	xInit			: BOOL;
	diPosPrev		: DINT;
	diTargetPrev	: DINT;
	diMoveStart		: DINT;

	xDirRev			: BOOL;
	xNewMove		: BOOL;
	xMoveWanted		: BOOL;
	xBrakeOpen		: BOOL;
	xMoving			: BOOL;
	xRunPrev		: BOOL;

	diStopAccum		: DINT;
	xCoasting		: BOOL;

	rtrgGo			: R_TRIG;
	rtrgReset		: R_TRIG;
	rtrgSetAccum	: R_TRIG;

	tofBrake		: TOF;
	tonBrakeOpen	: TON;
	tonGrace		: TON;
	tonStall		: TON;
	tonRest			: TON;
	tonDrvAck		: TON;

	diStallRef		: DINT;
	xStallReset		: BOOL;
	xStallArmed		: BOOL;

END_VAR

// =============================================================
// ENKODER -> PRZYROST ZE ZNAKIEM
// =============================================================
//
// Surowa wartosc moze byc wieksza niz jeden obrot, wiec
// sprowadzamy ja modulo. MOD na ujemnej daje w ST wynik ujemny,
// dlatego domykamy recznie.

diPos := diRawPos MOD 65536;

IF diPos < 0 THEN
	diPos := diPos + 65536;
END_IF


IF NOT xInit THEN
	xInit        := TRUE;
	diPosPrev    := diPos;
	diStallRef   := diPos;
	diTargetPrev := diTargetAbs;
END_IF


// Skok wiekszy niz pol obrotu nie jest ruchem - to licznik
// przekrecil sie przez zero. Prostujemy go i liczymy przejscie.

diStep := diPos - diPosPrev;

IF diStep > 32768 THEN
	diStep  := diStep - 65536;
	diTurns := diTurns - 1;
END_IF

IF diStep < -32768 THEN
	diStep  := diStep + 65536;
	diTurns := diTurns + 1;
END_IF

diPosPrev := diPos;


// =============================================================
// POZYCJA NARASTAJACA
// =============================================================
//
// Tu przestaje istniec problem przekrecania sie enkodera.
// diAccum jest zwykla liczba impulsow od punktu odniesienia
// i rosnie miedzy obrotami bez zadnego zawijania.

diAccum := diAccum + diStep;


// Punkt odniesienia ustawiany z zewnatrz, raz na cykl
rtrgSetAccum(CLK := xSetAccum);

IF rtrgSetAccum.Q THEN
	diAccum     := diSetAccumTo;
	diMoveStart := diSetAccumTo;
	xInPos      := TRUE;

	// Pomiar dojazdu musi przejsc przez ten skok sucha stopa.
	// diCoast liczy sie jako roznica na skali narastajacej,
	// wiec przestawienie punktu odniesienia bez tego wygladalo
	// by jak dojazd o caly obrot.
	diStopAccum := diSetAccumTo;
	xCoasting   := FALSE;
END_IF


// =============================================================
// NOWY RUCH
// =============================================================
//
// Nowy ruch to podanie zadania albo zmiana celu. diTargetAbs
// ma byc STALA w obrebie kroku - inaczej kazdy cykl wygladalby
// jak nowy ruch.

rtrgGo(CLK := xGoTo AND xEnable);

xNewMove := rtrgGo.Q OR (diTargetAbs <> diTargetPrev);
diTargetPrev := diTargetAbs;

IF xNewMove THEN
	diMoveStart := diAccum;
	xInPos      := FALSE;
	diStallRef  := diPos;
END_IF


// =============================================================
// UCHYB I KONIEC RUCHU
// =============================================================
//
// Zwykle odejmowanie, bez modulo. Uchyb ujemny znaczy "cel juz
// przejechany" i konczy ruch NATYCHMIAST - to jest dokladnie
// ten przypadek, w ktorym stara wersja wysylala os na dodatkowy
// pelen obrot.
//
// xInPos jest zatrzaskiem: osuniecie sie wozka po zacisnieciu
// hamulca nie ma prawa odwolac zaliczonego kroku.

diRemain := diTargetAbs - diAccum;
diMoved  := diAccum - diMoveStart;

IF diRemain <= diStopLead THEN
	xInPos := TRUE;
END_IF


// =============================================================
// RUCH I HAMULEC
// =============================================================
//
// Hamulec idzie za ZADANIEM ruchu, falownik dostaje komende
// tBrakeReleaseLead pozniej. Przy zerze - jednoczesnie.

xJogging := xEnable AND (xJogFwd XOR xJogRev);

xMoveWanted := xEnable AND NOT xStall AND (xJogging OR (xGoTo AND NOT xInPos));

// W cyklu korba jedzie WYLACZNIE do przodu. Kierunek wymuszamy
// co cykl, zeby ten z jazdy recznej w tyl nie mogl przezyc.
xDirRev := FALSE;

IF xJogging THEN
	xDirRev := xJogRev;
END_IF


tofBrake(IN := xMoveWanted, PT := tBrakeHold);
xBrakeRelease := tofBrake.Q;

tonBrakeOpen(IN := xMoveWanted AND xBrakeRelease, PT := tBrakeReleaseLead);

// Warunek na zero jawny - nie opieramy sie na tym, jak TON
// zachowa sie przy PT = 0. Blad w te strone dalby os, ktora
// nigdy nie rusza, i nic by tego nie powiedzialo.
xBrakeOpen := tonBrakeOpen.Q OR (tBrakeReleaseLead = T#0S);

xBrakeWait := xMoveWanted AND NOT xBrakeOpen;

xMoving := xMoveWanted AND xBrakeRelease AND xBrakeOpen;

xRunReq := xMoving;
xRev    := xDirRev;


// =============================================================
// POMIAR DOJAZDU
// =============================================================

IF xRunPrev AND NOT xRunReq THEN
	diStopAccum := diAccum;
	xCoasting   := TRUE;
END_IF

xRunPrev := xRunReq;

IF xCoasting THEN
	diCoast := diAccum - diStopAccum;
END_IF

tonRest(IN := ABS(diStep) < diStallMin, PT := tRest);
xAtRest := tonRest.Q;

IF xAtRest THEN
	xCoasting := FALSE;
END_IF


// =============================================================
// CZUWAK RUCHU
// =============================================================
//
// Uzbrojony dopiero po tStallGrace od startu - hamulec musi
// odpuscic, a silnik rozbiec sie rampa.

tonGrace(IN := xRunReq, PT := tStallGrace);
xStallArmed := tonGrace.Q;

xStallReset := (ABS(diAccum - diStallRef) > diStallMin)
               OR NOT xStallArmed OR xNewMove;

IF xStallReset THEN
	diStallRef := diAccum;
END_IF

tonStall(IN := xStallArmed AND NOT xStallReset, PT := tStall);

IF tonStall.Q THEN
	xStall := TRUE;
END_IF


// -------------------------------------------------------------
// POTWIERDZENIE PRACY Z FALOWNIKA
// -------------------------------------------------------------
//
// Osobny, szybszy czuwak. Zadanie poszlo, hamulec zdjety,
// a falownik nie melduje pracy - nic nie trzyma wozka i nie ma
// na co czekac pelnych pieciu sekund.

tonDrvAck(IN := xRunReq AND NOT xDrvRunning, PT := tDrvAck);

IF tonDrvAck.Q THEN
	xNoDrvAck := TRUE;
	xStall    := TRUE;
END_IF


rtrgReset(CLK := xReset);

IF rtrgReset.Q OR NOT xEnable THEN
	xStall     := FALSE;
	xNoDrvAck  := FALSE;
	diStallRef := diAccum;
END_IF

END_FUNCTION_BLOCK

// ---- POUs/POUs/FB/FB_NordSK550PP.TcPOU
FUNCTION_BLOCK FB_NordSK550PP
// =============================================================
// NORDAC PRO SK 550P
// EtherCAT, profil NORD wg BU 2300 (NIE CiA 402)
// =============================================================
//
// FB nie wykonuje ZADNYCH operacji na predkosci.
// Zadanie jest podawane na stale, sterowanie odbywa sie
// wylacznie bitami ControlWord. Rozpedzanie i hamowanie
// realizuje falownik parametrami P102 / P103 / P108.
//
// Sterowanie przez metody:
//   M_Start(lrFreq, xReverse)   - zadanie + bit startu
//   M_Stop()                    - zdjecie bitu startu
//   M_Reset()                   - kasowanie bledow
//   M_SetFrequency(lrFreq)      - zmiana zadania
//
// Metody wywolywac PRZED cyklicznym wywolaniem instancji.
VAR_INPUT

	// P105 Maksymalna czestotliwosc falownika [Hz].
	// MUSI byc rowna P105 w falowniku - inaczej skalowanie
	// zadania jest bledne i naped dostaje inna czestotliwosc
	// niz zadana.
	lrFmax			: LREAL := 50.0;

	// TRUE = STO zwolnione, lancuch bezpieczenstwa OK
	xSafetyOK		: BOOL;

	// TRUE = komunikacja EtherCAT sprawna
	xEtherCAT_OK	: BOOL;

	// Dane procesowe z falownika
	stIn			: ST_NordSK550P_In;

END_VAR
VAR_OUTPUT

	// Dane procesowe do falownika
	stOut			: ST_NordSK550P_Out;


	// =========================================================
	// STATUS
	// =========================================================

	eState			: E_NordSK550P_State;

	xReadyToSwitchOn	: BOOL;
	xOperationEnabled	: BOOL;
	xSwitchOnInhibit	: BOOL;

	xRunning		: BOOL;
	xStopped		: BOOL;

	xFault			: BOOL;
	xWarning		: BOOL;
	xBusControl		: BOOL;

	xError			: BOOL;
	xCommError		: BOOL;


	// =========================================================
	// VALUES
	// =========================================================

	// Zadanie wysylane do falownika [Hz]
	lrFreqSetpoint	: LREAL;

	// Czestotliwosc rzeczywista z falownika [Hz]
	lrFreqActual	: LREAL;


	// =========================================================
	// DIAGNOSTICS
	// =========================================================

	wStatusWord		: UINT;
	wControlWord	: UINT;

	byModeDisplay	: USINT;

	//  0 = blokada, 10 = gotowosc, 20 = praca
	nStep			: INT;

END_VAR
VAR

	// Zadania z metod
	xReqRun			: BOOL;
	xReqReset		: BOOL;
	xReqReverse		: BOOL;
	lrReqFreq		: LREAL;

	wStateBits		: UINT;
	iSetpoint		: INT;
	xBlocked		: BOOL;

	tonComm			: TON;
	tonReset		: TON;

END_VAR
VAR CONSTANT

	// Skalowanie NORD: 16384 (0x4000) = 100% = P105
	cFullScale		: LREAL := 16384.0;

	// Prog zera dla czestotliwosci rzeczywistej [Hz]
	cZeroActual		: LREAL := 0.5;

	// ControlWord wg BU 2300 rozdz. 6.3.1
	//   047E = "Shut down"        - bit 0 zdjety, falownik
	//                               hamuje wlasna rampa P103
	//   047F = "Enable operation" - bit 0 zalaczony
	//   0480 = potwierdzenie bledu (bit 7)
	cCW_Shutdown	: UINT := 16#047E;
	cCW_EnableOp	: UINT := 16#047F;
	cCW_AckFault	: UINT := 16#0480;

	cCW_DirFwd		: UINT := 16#0800;
	cCW_DirRev		: UINT := 16#1000;

END_VAR

// =============================================================
// FB_NordSK550PP
// NORDAC PRO SK 550P - profil NORD wg BU 2300
// =============================================================
//
// ZASADA: PLC nie dotyka predkosci.
//
// Zadanie czestotliwosci jest podawane na stale i nie jest
// zerowane przy zatrzymaniu. Start to zalaczenie bitu 0
// ControlWord, stop to jego zdjecie. Reszte - rozpedzanie
// po P102, hamowanie po P103, sposob wygaszania po P108
// i ewentualne dohamowanie pradem stalym po P559 - robi
// falownik.
//
// ControlWord (BU 2300 rozdz. 6.3.1):
//   bit 0  Ready for operation   <-- start / stop
//   bit 1  Voltage disable       (1 = kasuj blokade napiecia)
//   bit 2  Quick stop            (1 = kasuj quick stop)
//   bit 3  Enable operation
//   bit 4  Enable pulses
//   bit 5  Enable ramp
//   bit 6  Setpoint enabled
//   bit 7  Acknowledge error     (zbocze 0 -> 1)
//   bit 10 Control data valid    <-- BEZ NIEGO NAPED IGNORUJE DANE
//   bit 11 CW, bit 12 CCW
//
// StatusWord (rozdz. 6.3.2), bity 0..6:
//   0x31 Ready to switch-on   0x33 Switched on
//   0x37 Operation enabled    0x17 Quick stop active
//   bit 3 Fault               bit 6 Switch-on inhibit
//
// Zadanie i wartosc rzeczywista sa procentowe:
//   16384 (0x4000) = 100% = P105
//
// Nazwy pol diTargetVelocity / iVelocityDemand w ST_NordSK550P_*
// sa mylace - to NIE obroty, tylko czestotliwosc w skali
// procentowej. NIE zmieniac tych nazw: sa uzyte w linkach I/O
// w .tsproj dla wszystkich 19 napedow.


// =============================================================
// COPY INPUT DATA
// =============================================================

wStatusWord		:= stIn.wStatusWord;
byModeDisplay	:= stIn.byModeDisplay;

IF lrFmax > 0.0 THEN
	lrFreqActual := INT_TO_LREAL(stIn.iVelocityDemand) / cFullScale * lrFmax;
ELSE
	lrFreqActual := 0.0;
END_IF


// =============================================================
// COMMUNICATION WATCHDOG
// =============================================================

tonComm(IN := NOT xEtherCAT_OK, PT := T#500MS);
xCommError := tonComm.Q;


// =============================================================
// STATUSWORD DECODING
// =============================================================

xFault				:= (wStatusWord AND 16#0008) <> 0;
xWarning			:= (wStatusWord AND 16#0080) <> 0;
xSwitchOnInhibit	:= (wStatusWord AND 16#0040) <> 0;
xBusControl			:= (wStatusWord AND 16#0200) <> 0;

wStateBits := wStatusWord AND 16#007F;


IF xFault THEN

	IF (wStatusWord AND 16#000F) = 16#000F THEN
		eState := NORD_STATE_FAULT_REACTION_ACTIVE;
	ELSE
		eState := NORD_STATE_FAULT;
	END_IF

ELSIF xSwitchOnInhibit THEN
	eState := NORD_STATE_SWITCH_ON_DISABLED;

ELSIF wStateBits = 16#0031 THEN
	eState := NORD_STATE_READY_TO_SWITCH_ON;

ELSIF wStateBits = 16#0033 THEN
	eState := NORD_STATE_SWITCHED_ON;

ELSIF wStateBits = 16#0037 THEN
	eState := NORD_STATE_OPERATION_ENABLED;

ELSIF wStateBits = 16#0017 THEN
	eState := NORD_STATE_QUICK_STOP_ACTIVE;

ELSIF (wStatusWord AND 16#000F) = 0 THEN
	eState := NORD_STATE_NOT_READY;

ELSE
	eState := NORD_STATE_UNKNOWN;

END_IF


xReadyToSwitchOn	:= (eState = NORD_STATE_READY_TO_SWITCH_ON);
xOperationEnabled	:= (eState = NORD_STATE_OPERATION_ENABLED);


// =============================================================
// WARUNKI BLOKUJACE
// =============================================================

xBlocked := xFault OR xCommError OR NOT xSafetyOK;
xError   := xBlocked;


// =============================================================
// CONTROLWORD
// =============================================================
//
// Trzy stany, bez zadnej sekwencji posredniej. Przejscia
// wewnetrznej maszyny stanow falownika (Switch-on inhibit ->
// Ready to switch-on -> Switched on -> Operation enabled)
// realizuje sam falownik: 047E zawiera komende "Shut down",
// a 047F jednoczesnie "Switch on" i "Enable operation".

IF xBlocked THEN

	nStep := 0;

	// Zadanie ruchu kasujemy - po ustapieniu przyczyny naped
	// NIE moze ruszyc sam, operator musi wywolac M_Start.
	xReqRun := FALSE;

	wControlWord := 16#0000;

	// Kasowanie bledu: impuls na bicie 7
	IF xReqReset AND xSafetyOK AND NOT xCommError THEN
		wControlWord := cCW_AckFault;
	END_IF

ELSIF xReqRun THEN

	nStep := 20;
	wControlWord := cCW_EnableOp;

	// BLOKADA ZALACZENIA (Switch-on inhibit, bit 6 statusu).
	//
	// Ze stanu "Switch on disabled" falownik NIE wyjdzie na 047F.
	// Bit 0 musi zobaczyc zbocze, a zeby je zobaczyl, trzeba
	// najpierw wyslac Shutdown (047E). Trzymanie 047F w kolko
	// zostawia naped w blokadzie na zawsze: bez bledu, bez ruchu,
	// bez zadnego komunikatu - dokladnie to widzielismy na
	// napedzie 5 po przeciazeniu i na 8 po zaniku komunikacji.
	//
	// Dopoki falownik melduje blokade, wysylamy wiec 047E. Gdy
	// z niej wyjdzie, w nastepnym cyklu idzie juz 047F i naped
	// rusza sam, bez kasowania bledu i bez zdejmowania startu.
	IF xSwitchOnInhibit THEN
		nStep := 15;
		wControlWord := cCW_Shutdown;
	END_IF

ELSE

	nStep := 10;
	wControlWord := cCW_Shutdown;

END_IF


// =============================================================
// KIERUNEK
// =============================================================
//
// Zmiane kierunku w ruchu obsluguje falownik - przechodzi
// przez absolutna minimalna czestotliwosc P505.

IF wControlWord <> 16#0000 THEN

	IF xReqReverse THEN
		wControlWord := wControlWord OR cCW_DirRev;
	ELSE
		wControlWord := wControlWord OR cCW_DirFwd;
	END_IF

END_IF


// =============================================================
// IMPULS KASOWANIA BLEDU
// =============================================================
//
// Bit 7 musi zobaczyc zbocze 0 -> 1. Trzymamy go 200 ms,
// potem kasujemy zadanie, zeby kolejne M_Reset znowu
// wytworzylo zbocze.

tonReset(IN := xReqReset, PT := T#200MS);

IF tonReset.Q THEN
	xReqReset := FALSE;
END_IF


// =============================================================
// ZADANIE CZESTOTLIWOSCI
// =============================================================
//
// Podawane na stale. NIE zerujemy go przy zatrzymaniu -
// stop realizuje bit 0 ControlWord, a hamowanie falownik.

lrFreqSetpoint := lrReqFreq;

IF lrFreqSetpoint > lrFmax THEN
	lrFreqSetpoint := lrFmax;
END_IF

IF lrFreqSetpoint < 0.0 THEN
	lrFreqSetpoint := 0.0;
END_IF


IF lrFmax > 0.0 THEN
	iSetpoint := LREAL_TO_INT(lrFreqSetpoint / lrFmax * cFullScale);
ELSE
	iSetpoint := 0;
END_IF

IF iSetpoint > 16384 THEN
	iSetpoint := 16384;
END_IF

IF iSetpoint < 0 THEN
	iSetpoint := 0;
END_IF


// =============================================================
// WRITE OUTPUT PDO
// =============================================================
//
// byModeOfOperation nie jest zmapowany w .tsproj - falownik
// NORD nie uzywa obiektu 0x6060. Zostawiamy zero.

stOut.byModeOfOperation	:= 0;
stOut.wControlWord		:= wControlWord;
stOut.diTargetVelocity	:= iSetpoint;


// =============================================================
// STATUS WYJSCIOWY
// =============================================================

xRunning := xOperationEnabled AND NOT xBlocked;

xStopped := (ABS(lrFreqActual) <= cZeroActual);

METHOD M_Start : BOOL
VAR_INPUT
	// Zadana czestotliwosc [Hz]
	lrFreq		: LREAL;

	// FALSE = w prawo (CW), TRUE = w lewo (CCW)
	xReverse	: BOOL;
END_VAR
// Zadanie czestotliwosci + bit startu. Nic wiecej.
// Rozpedzanie realizuje falownik rampa P102.
//
// Zadanie jest zatrzaskiwane - obowiazuje az do M_Stop
// albo do wystapienia blokady (blad / STO / komunikacja).

lrReqFreq	:= lrFreq;
xReqReverse	:= xReverse;
xReqRun		:= TRUE;

M_Start := TRUE;
END_METHOD

METHOD M_Stop : BOOL
// Zdjecie bitu 0 ControlWord. Nic wiecej - zadanie
// czestotliwosci zostaje bez zmian.
//
// Falownik hamuje wlasna rampa P103, sposob wygaszania
// okresla P108, ewentualne dohamowanie pradem stalym P559.

xReqRun := FALSE;

M_Stop := TRUE;
END_METHOD

METHOD M_Reset : BOOL
// Kasowanie bledow falownika. FB wystawia impuls 200 ms
// na bicie 7 ControlWord (zbocze 0 -> 1 wg BU 2300).
//
// Dziala tylko wtedy, gdy przyczyna blokady ustapila:
// STO zwolnione i komunikacja sprawna.

xReqReset := TRUE;

M_Reset := TRUE;
END_METHOD

METHOD M_SetFrequency : BOOL
VAR_INPUT
	// Zadana czestotliwosc [Hz]
	lrFreq		: LREAL;
END_VAR
// Zmiana zadania. Falownik dojezdza do nowej wartosci
// wlasna rampa.

lrReqFreq := lrFreq;

M_SetFrequency := TRUE;
END_METHOD

END_FUNCTION_BLOCK

// ---- POUs/POUs/FB/FB_CsvLogger.TcPOU
FUNCTION_BLOCK FB_CsvLogger
// =============================================================
// OBSERWATOR STANU MASZYNY - ZAPIS CSV NA DYSK STEROWNIKA
// =============================================================
//
// Blok NICZEGO nie zapisuje do zmiennych procesu. Tylko czyta
// to, co mu poda MAIN, i odklada na dysk.
//
// -------------------------------------------------------------
// JAK SIE TEGO UZYWA (ACT_Logger w MAIN)
// -------------------------------------------------------------
//
//   fbLog.M_Begin();
//   fbLog.M_Int ('nDeStep', nDeStep);
//   fbLog.M_Bool('xPal_St03', xPal_St03);
//   ...
//   fbLog.M_End();
//
// Kazda metoda M_* dostaje NAZWE kolumny i WARTOSC. Gdy
// xHeaderMode = TRUE, metoda dopisuje nazwe zamiast wartosci -
// dzieki temu naglowek i wiersz powstaja z tego samego kodu
// i nie moga sie rozjechac.
//
// -------------------------------------------------------------
// PLIK
// -------------------------------------------------------------
//
// Nazwa: <sDir><sPrefix>_RRRRMMDD_GGMMSS.csv, czas z zegara
// sterownika (NT_GetTime). Nowy plik na zbocze xNewFile.
//
// Kazdy zrzut to OTWORZ (append) -> ZAPISZ -> ZAMKNIJ. Uchwyt
// nie jest trzymany miedzy zrzutami, wiec:
//   - plik mozna kopiowac w trakcie pracy,
//   - stop PLC nie gubi ostatniego bufora,
//   - katalog zaklada FB_CreateDir przy pierwszym starcie;
//     jesli sie nie uda, nMkDirErrId to pokaze.
//
// Wiersze zbieraja sie w kolejce aOut i ida na dysk jednym
// zapisem, nie czesciej niz co tFlushMin. Operacje na pliku sa
// asynchroniczne (ADS) - cykl PLC na dysk nigdy nie czeka.
//
// Gdy kolejka jest pelna, wiersz przepada i rosnie
// nLinesDropped. Lepiej zgubic wiersz niz cykl.
VAR_INPUT

	// Katalog z koncowym ukosnikiem. Zakladany automatycznie.
	sDir			: STRING(200) := 'C:\TesterPalet\log\';

	// Poczatek nazwy pliku
	sPrefix			: STRING(31) := 'tp';

	// Zbocze 0 -> 1 = zamknij biezacy plik, zaloz nowy
	xNewFile		: BOOL;

	// Najkrotszy odstep miedzy zrzutami na dysk
	tFlushMin		: TIME := T#500MS;

	// Limit czasu jednej operacji ADS na pliku
	tTimeout		: TIME := T#3S;

	// TRUE = metody M_* dopisuja NAZWE kolumny, nie wartosc
	xHeaderMode		: BOOL;

END_VAR
VAR_OUTPUT

	// Nazwa biezacego pliku - do odczytu online
	sFileName		: STRING(255);

	// TRUE = plik nazwany, ale naglowek jeszcze nie poszedl.
	// MAIN na tym bicie wysyla wiersz naglowka.
	xHeaderPending	: BOOL;

	// Milisekundy od otwarcia pliku - kolumna t_ms
	udiFileMs		: UDINT;

	// Statystyka
	nFileNo			: UDINT;
	nLinesQueued	: UDINT;
	nLinesDropped	: UDINT;
	nBytesWritten	: UDINT;
	nFlushes		: UDINT;
	nErrors			: UDINT;
	nLastErrId		: UDINT;
	sLastErrWhere	: STRING(15);

	// Podglad maszyny stanu bloku
	nState			: INT;

	// Wynik zakladania katalogu: 0 = OK albo juz istnial
	nMkDirErrId		: UDINT;

	// Bajty czekajace w kolejce
	nOutLen			: UDINT;

END_VAR
VAR

	xInit			: BOOL;
	xRotateReq		: BOOL;
	xFileNamed		: BOOL;
	xFlushTick		: BOOL;

	// Skladany wiersz
	aLine			: ARRAY[0..cLineMax] OF BYTE;
	nLineLen		: UDINT;
	xLineOverflow	: BOOL;

	// Kolejka wierszy czekajacych na zrzut
	aOut			: ARRAY[0..cOutMax] OF BYTE;

	// Bufor w trakcie zapisu - FB_FileWrite trzyma wskaznik,
	// wiec kolejka nie moze sie pod nim zmieniac
	aWr				: ARRAY[0..cOutMax] OF BYTE;
	nWrLen			: UDINT;

	fbOpen			: FB_FileOpen;
	fbWrite			: FB_FileWrite;
	fbClose			: FB_FileClose;
	fbTime			: NT_GetTime;		// Tc2_Utilities
	fbMkDir			: FB_CreateDir;		// Tc2_Utilities
	hFile			: UINT;
	xDirDone		: BOOL;
	sDirNoSlash		: STRING(200);

	rtrgNew			: R_TRIG;
	tonFlush		: TON;

	// Zegar: milisekundy doby w chwili otwarcia pliku
	udiStartMsOfDay	: UDINT;
	tFileStart		: TIME;

	// Robocze
	sTmp			: STRING(63);
	nTmp			: DINT;

END_VAR
VAR CONSTANT

	cLineMax		: UDINT := 8191;
	cOutMax			: UDINT := 65535;
	cCR				: BYTE := 13;
	cLF				: BYTE := 10;
	cSep			: BYTE := 59;		// ';'

END_VAR

// =============================================================
// ZBOCZE NOWEGO PLIKU
// =============================================================

rtrgNew(CLK := xNewFile);

IF rtrgNew.Q OR NOT xInit THEN
	xInit      := TRUE;
	xRotateReq := TRUE;
END_IF


// Takt zrzutu - nie czesciej niz tFlushMin
tonFlush(IN := TRUE, PT := tFlushMin);
xFlushTick := tonFlush.Q;

IF xFlushTick THEN
	tonFlush(IN := FALSE);
END_IF


// Milisekundy od otwarcia pliku
IF xFileNamed THEN
	udiFileMs := TIME_TO_UDINT(TIME() - tFileStart);
END_IF


// =============================================================
// MASZYNA STANU ZAPISU
// =============================================================
//
//   0   spokoj: czekam na zrzut albo na nowy plik
//   5   zakladam katalog (raz, przy pierwszym starcie)
//  10   pobieram czas z zegara sterownika -> nazwa pliku
//  20   otwieram plik (append)
//  30   pisze bufor aWr
//  40   zamykam plik

CASE nState OF

0:
	IF xRotateReq AND NOT xDirDone THEN
		// Katalog bez koncowego ukosnika
		sDirNoSlash := sDir;
		IF RIGHT(sDirNoSlash, 1) = '\' THEN
			sDirNoSlash := LEFT(sDirNoSlash, LEN(sDirNoSlash) - 1);
		END_IF
		fbMkDir(bExecute := FALSE);
		nState := 5;
	ELSIF xRotateReq THEN
		xRotateReq := FALSE;
		fbTime(NETID := '', START := FALSE);
		nState := 10;
	ELSIF xFileNamed AND (nOutLen > 0) AND xFlushTick THEN
		MEMCPY(destAddr := ADR(aWr), srcAddr := ADR(aOut), n := nOutLen);
		nWrLen  := nOutLen;
		nOutLen := 0;
		fbOpen(bExecute := FALSE);
		nState := 20;
	END_IF

5:
	fbMkDir(
		sNetId    := '',
		sPathName := sDirNoSlash,
		ePath     := PATH_GENERIC,
		bExecute  := TRUE,
		tTimeout  := tTimeout);

	IF NOT fbMkDir.bBusy THEN
		// Blad "juz istnieje" jest w porzadku - tylko do podgladu
		nMkDirErrId := 0;
		IF fbMkDir.bError THEN
			nMkDirErrId := fbMkDir.nErrId;
		END_IF
		fbMkDir(bExecute := FALSE);
		xDirDone := TRUE;
		nState   := 0;
	END_IF

10:
	fbTime(NETID := '', START := TRUE, TMOUT := tTimeout);

	IF NOT fbTime.BUSY THEN

		nFileNo := nFileNo + 1;

		IF fbTime.ERR THEN
			// Bez zegara tez logujemy - nazwa z licznika
			sFileName := CONCAT(sDir, sPrefix);
			sFileName := CONCAT(sFileName, '_noclock_');
			sFileName := CONCAT(sFileName, UDINT_TO_STRING(nFileNo));
			sFileName := CONCAT(sFileName, '.csv');
			udiStartMsOfDay := 0;
			nErrors    := nErrors + 1;
			nLastErrId := fbTime.ERRID;
			sLastErrWhere := 'NT_GetTime';
		ELSE
			sFileName := CONCAT(sDir, sPrefix);
			sFileName := CONCAT(sFileName, '_');
			sFileName := CONCAT(sFileName, WORD_TO_STRING(fbTime.TIMESTR.wYear));
			sFileName := CONCAT(sFileName, M_Pad2(fbTime.TIMESTR.wMonth));
			sFileName := CONCAT(sFileName, M_Pad2(fbTime.TIMESTR.wDay));
			sFileName := CONCAT(sFileName, '_');
			sFileName := CONCAT(sFileName, M_Pad2(fbTime.TIMESTR.wHour));
			sFileName := CONCAT(sFileName, M_Pad2(fbTime.TIMESTR.wMinute));
			sFileName := CONCAT(sFileName, M_Pad2(fbTime.TIMESTR.wSecond));
			sFileName := CONCAT(sFileName, '.csv');
			udiStartMsOfDay := WORD_TO_UDINT(fbTime.TIMESTR.wHour) * 3600000
			                 + WORD_TO_UDINT(fbTime.TIMESTR.wMinute) * 60000
			                 + WORD_TO_UDINT(fbTime.TIMESTR.wSecond) * 1000
			                 + WORD_TO_UDINT(fbTime.TIMESTR.wMilliseconds);
		END_IF

		fbTime(NETID := '', START := FALSE);

		tFileStart     := TIME();
		udiFileMs      := 0;
		xFileNamed     := TRUE;
		xHeaderPending := TRUE;
		nState         := 0;
	END_IF

20:
	fbOpen(
		sNetId    := '',
		sPathName := sFileName,
		nMode     := FOPEN_MODEAPPEND OR FOPEN_MODEBINARY,
		ePath     := PATH_GENERIC,
		bExecute  := TRUE,
		tTimeout  := tTimeout);

	IF NOT fbOpen.bBusy THEN
		IF fbOpen.bError THEN
			nErrors       := nErrors + 1;
			nLastErrId    := fbOpen.nErrId;
			sLastErrWhere := 'FB_FileOpen';
			fbOpen(bExecute := FALSE);
			nState := 0;
		ELSE
			hFile := fbOpen.hFile;
			fbWrite(bExecute := FALSE);
			nState := 30;
		END_IF
	END_IF

30:
	fbWrite(
		sNetId     := '',
		hFile      := hFile,
		pWriteBuff := ADR(aWr),
		cbWriteLen := nWrLen,
		bExecute   := TRUE,
		tTimeout   := tTimeout);

	IF NOT fbWrite.bBusy THEN
		IF fbWrite.bError THEN
			nErrors       := nErrors + 1;
			nLastErrId    := fbWrite.nErrId;
			sLastErrWhere := 'FB_FileWrite';
		ELSE
			nBytesWritten := nBytesWritten + fbWrite.cbWrite;
			nFlushes      := nFlushes + 1;
		END_IF
		fbWrite(bExecute := FALSE);
		fbClose(bExecute := FALSE);
		nState := 40;
	END_IF

40:
	fbClose(
		sNetId   := '',
		hFile    := hFile,
		bExecute := TRUE,
		tTimeout := tTimeout);

	IF NOT fbClose.bBusy THEN
		IF fbClose.bError THEN
			nErrors       := nErrors + 1;
			nLastErrId    := fbClose.nErrId;
			sLastErrWhere := 'FB_FileClose';
		END_IF
		fbClose(bExecute := FALSE);
		fbOpen(bExecute := FALSE);
		nState := 0;
	END_IF

ELSE
	nState := 0;

END_CASE

// Poczatek wiersza - czysci bufor skladania
METHOD M_Begin
nLineLen      := 0;
xLineOverflow := FALSE;
END_METHOD

// Koniec wiersza - CRLF i do kolejki.
// Naglowek (xHeaderMode) idzie na POCZATEK kolejki, zeby byl
// pierwsza linia pliku nawet wtedy, gdy wiersze zdazyly sie
// juz ustawic w kolejce przed nadaniem nazwy.
METHOD M_End
VAR
	nNeed	: UDINT;
END_VAR
IF nLineLen = 0 THEN
	RETURN;
END_IF

// Ostatni srednik zamieniamy na koniec linii
IF aLine[nLineLen - 1] = cSep THEN
	nLineLen := nLineLen - 1;
END_IF

IF nLineLen + 2 > cLineMax THEN
	xLineOverflow := TRUE;
END_IF

IF xLineOverflow THEN
	nLinesDropped := nLinesDropped + 1;
	nLineLen := 0;
	RETURN;
END_IF

aLine[nLineLen]     := cCR;
aLine[nLineLen + 1] := cLF;
nNeed := nLineLen + 2;

IF nOutLen + nNeed > cOutMax THEN
	nLinesDropped := nLinesDropped + 1;
	nLineLen := 0;
	RETURN;
END_IF

IF xHeaderMode THEN
	IF nOutLen > 0 THEN
		MEMMOVE(destAddr := ADR(aOut[nNeed]), srcAddr := ADR(aOut), n := nOutLen);
	END_IF
	MEMCPY(destAddr := ADR(aOut), srcAddr := ADR(aLine), n := nNeed);
	xHeaderPending := FALSE;
ELSE
	MEMCPY(destAddr := ADR(aOut[nOutLen]), srcAddr := ADR(aLine), n := nNeed);
END_IF

nOutLen      := nOutLen + nNeed;
nLinesQueued := nLinesQueued + 1;
nLineLen     := 0;
END_METHOD

// Dopisz tekst do wiersza BEZ separatora. Sredniki w tresci
// zamienia na przecinki, zeby nie rozbily kolumn.
METHOD M_Raw
VAR_INPUT
	sText	: STRING(255);
END_VAR
VAR
	nLen	: UDINT;
	i		: UDINT;
	pByte	: POINTER TO BYTE;
END_VAR
nLen := INT_TO_UDINT(LEN(sText));

IF nLen = 0 THEN
	RETURN;
END_IF

IF nLineLen + nLen > cLineMax THEN
	xLineOverflow := TRUE;
	RETURN;
END_IF

MEMCPY(destAddr := ADR(aLine[nLineLen]), srcAddr := ADR(sText), n := nLen);

pByte := ADR(aLine[nLineLen]);

FOR i := 0 TO nLen - 1 DO
	IF pByte^ = cSep THEN
		pByte^ := 44;	// ','
	END_IF
	IF pByte^ < 32 THEN
		pByte^ := 32;	// znaki sterujace -> spacja
	END_IF
	pByte := pByte + 1;
END_FOR

nLineLen := nLineLen + nLen;
END_METHOD

// Separator kolumn
METHOD M_Sep
IF nLineLen + 1 > cLineMax THEN
	xLineOverflow := TRUE;
	RETURN;
END_IF

aLine[nLineLen] := cSep;
nLineLen := nLineLen + 1;
END_METHOD

// Kolumna tekstowa
METHOD M_Str
VAR_INPUT
	sName	: STRING(63);
	sVal	: STRING(255);
END_VAR
IF xHeaderMode THEN
	M_Raw(sName);
ELSE
	M_Raw(sVal);
END_IF

M_Sep();
END_METHOD

// Kolumna calkowita (INT, DINT, UDINT po konwersji)
METHOD M_Int
VAR_INPUT
	sName	: STRING(63);
	diVal	: DINT;
END_VAR
IF xHeaderMode THEN
	M_Raw(sName);
ELSE
	M_Raw(DINT_TO_STRING(diVal));
END_IF

M_Sep();
END_METHOD

// Kolumna calkowita bez znaku (UDINT - liczniki)
METHOD M_UInt
VAR_INPUT
	sName	: STRING(63);
	udiVal	: UDINT;
END_VAR
IF xHeaderMode THEN
	M_Raw(sName);
ELSE
	M_Raw(UDINT_TO_STRING(udiVal));
END_IF

M_Sep();
END_METHOD

// Kolumna logiczna: 1 / 0
METHOD M_Bool
VAR_INPUT
	sName	: STRING(63);
	xVal	: BOOL;
END_VAR
IF xHeaderMode THEN
	M_Raw(sName);
ELSIF xVal THEN
	M_Raw('1');
ELSE
	M_Raw('0');
END_IF

M_Sep();
END_METHOD

// Kolumna szesnastkowa 16-bit, np. 0637 (slowa stanu falownikow)
METHOD M_Hex
VAR_INPUT
	sName	: STRING(63);
	wVal	: WORD;
END_VAR
VAR
	aHex	: ARRAY[0..4] OF BYTE;
	sHex	: STRING(4);
	i		: INT;
	nNib	: BYTE;
END_VAR
IF xHeaderMode THEN
	M_Raw(sName);
ELSE
	FOR i := 0 TO 3 DO
		nNib := WORD_TO_BYTE(SHR(wVal, 12 - 4 * i) AND 16#000F);
		IF nNib < 10 THEN
			aHex[i] := 48 + nNib;		// '0'..'9'
		ELSE
			aHex[i] := 55 + nNib;		// 'A'..'F'
		END_IF
	END_FOR
	aHex[4] := 0;
	MEMCPY(destAddr := ADR(sHex), srcAddr := ADR(aHex), n := 5);
	M_Raw(sHex);
END_IF

M_Sep();
END_METHOD

// Kolumna zmiennoprzecinkowa z JEDNYM miejscem po kropce.
// LREAL_TO_STRING daje kilkanascie cyfr - nieczytelne w CSV.
METHOD M_Real
VAR_INPUT
	sName	: STRING(63);
	lrVal	: LREAL;
END_VAR
VAR
	diScaled	: DINT;
	diAbs		: DINT;
	sOut		: STRING(31);
END_VAR
IF xHeaderMode THEN
	M_Raw(sName);
ELSE
	diScaled := LREAL_TO_DINT(lrVal * 10.0);
	diAbs    := ABS(diScaled);
	sOut := DINT_TO_STRING(diAbs / 10);
	sOut := CONCAT(sOut, '.');
	sOut := CONCAT(sOut, DINT_TO_STRING(diAbs MOD 10));
	IF diScaled < 0 THEN
		sOut := CONCAT('-', sOut);
	END_IF
	M_Raw(sOut);
END_IF

M_Sep();
END_METHOD

// Kolumna zegara GG:MM:SS.mmm - czas otwarcia pliku plus
// milisekundy od otwarcia. Nie pyta zegara co cykl.
METHOD M_Clock
VAR_INPUT
	sName	: STRING(63);
END_VAR
VAR
	udiMs	: UDINT;
	sOut	: STRING(15);
END_VAR
IF xHeaderMode THEN
	M_Raw(sName);
ELSE
	udiMs := (udiStartMsOfDay + udiFileMs) MOD 86400000;
	sOut := M_Pad2(UDINT_TO_WORD(udiMs / 3600000));
	sOut := CONCAT(sOut, ':');
	sOut := CONCAT(sOut, M_Pad2(UDINT_TO_WORD((udiMs / 60000) MOD 60)));
	sOut := CONCAT(sOut, ':');
	sOut := CONCAT(sOut, M_Pad2(UDINT_TO_WORD((udiMs / 1000) MOD 60)));
	sOut := CONCAT(sOut, '.');
	sOut := CONCAT(sOut, M_Pad3(UDINT_TO_WORD(udiMs MOD 1000)));
	M_Raw(sOut);
END_IF

M_Sep();
END_METHOD

// Liczba 0..99 jako dwa znaki z zerem wiodacym
METHOD M_Pad2 : STRING(7)
VAR_INPUT
	wVal	: WORD;
END_VAR
IF wVal < 10 THEN
	M_Pad2 := CONCAT('0', WORD_TO_STRING(wVal));
ELSE
	M_Pad2 := WORD_TO_STRING(wVal);
END_IF
END_METHOD

// Liczba 0..999 jako trzy znaki z zerami wiodacymi
METHOD M_Pad3 : STRING(7)
VAR_INPUT
	wVal	: WORD;
END_VAR
IF wVal < 10 THEN
	M_Pad3 := CONCAT('00', WORD_TO_STRING(wVal));
ELSIF wVal < 100 THEN
	M_Pad3 := CONCAT('0', WORD_TO_STRING(wVal));
ELSE
	M_Pad3 := WORD_TO_STRING(wVal);
END_IF
END_METHOD

END_FUNCTION_BLOCK

// ---- POUs/POUs/FB/FB_StackLift.TcPOU
FUNCTION_BLOCK FB_StackLift
// =============================================================
// WOZEK ZE SZCZEKAMI - DESZTAPLARKA I SZTAPLARKA
// =============================================================
//
// Jedna kinematyka dla obu maszyn: wozek jezdzacy w pionie na
// falowniku NORD, enkoder absolutny i szczeki na siłowniku.
// Rozni je wylacznie kolejnosc krokow, ktora siedzi w stacjach.
//
// -------------------------------------------------------------
// TRZY POZYCJE
// -------------------------------------------------------------
//   POS_BOTTOM  deski pierwszej palety od dolu
//   POS_MIDDLE  deski drugiej palety od dolu
//   POS_TOP     stos uniesiony
//
// Odleglosc miedzy nimi to wysokosc palety - stad wszystkie trzy
// sa potrzebne i stad kontrola, ze tworza ciag. Wpisanie ich
// w zlej kolejnosci wyslaloby wozek w przeciwna strone niz
// trzeba, wiec sprawdzamy to, zanim ruszymy.
//
// -------------------------------------------------------------
// POZYCJONOWANIE
// -------------------------------------------------------------
// Falownik NORD dostaje wylacznie czestotliwosc, wiec dojazd
// jest dwustopniowy: pelna predkosc do strefy dojazdowej, potem
// predkosc dojazdowa do okna pozycji. Hamowanie realizuje rampa
// falownika (P103), tak jak wszedzie indziej w tym projekcie.
VAR_INPUT

	eMode			: E_MachineMode;
	xSafetyOK		: BOOL;

	// Enkoder absolutny wozka
	diPosRaw		: DINT;

	// Krancowki szczek - jesli ich nie ma, wylaczyc obserwacje
	// w rekordzie silownika i pracowac na czasowce
	xJawClosedSw	: BOOL;
	xJawOpenSw		: BOOL;

END_VAR
VAR_OUTPUT

	// Cewki szczek - stacja przepisuje na swoje wyjscia
	xJawCoilClose	: BOOL;
	xJawCoilOpen	: BOOL;

	diPos			: DINT;
	diTarget		: DINT;
	diError			: DINT;

	// 0 brak, 1 dol, 2 srodek, 3 gora
	nTargetSel		: INT;

	xInPosition		: BOOL;
	xMoving			: BOOL;
	xJawsClosed		: BOOL;
	xJawsOpen		: BOOL;

	eAlarm			: E_StackAlarm;
	xAlarm			: BOOL;

END_VAR
VAR

	pP				: POINTER TO ST_StackPersist;
	pDrive			: POINTER TO FB_NordSK550PP;

	fbJaw			: FB_Cylinder;

	xRunReq			: BOOL;
	xRevReq			: BOOL;
	lrFreqReq		: LREAL;

	xRunOld			: BOOL;
	xRevOld			: BOOL;
	lrFreqOld		: LREAL;

	tonMoveWd		: TON;
	tonSettle		: TON;

	xManUp			: BOOL;
	xManDown		: BOOL;

END_VAR

// =============================================================
// CYKL WOZKA
// =============================================================


// -------------------------------------------------------------
// 1. KONFIGURACJA
// -------------------------------------------------------------

IF pP = 0 THEN
	M_HaltDrive();
	eAlarm := ALM_STK_NOT_CONFIGURED;
	xAlarm := TRUE;
	RETURN;
END_IF

diPos	:= diPosRaw;
diError	:= diTarget - diPos;
xAlarm	:= (eAlarm <> ALM_STK_NONE);


// -------------------------------------------------------------
// 2. SZCZEKI
// -------------------------------------------------------------

fbJaw(
	eMode		:= eMode,
	xSafetyOK	:= xSafetyOK,
	xSwExtRaw	:= xJawClosedSw,
	xSwRetRaw	:= xJawOpenSw
);

xJawCoilClose	:= fbJaw.xCoilExtend;
xJawCoilOpen	:= fbJaw.xCoilRetract;
xJawsClosed		:= fbJaw.xExtended;
xJawsOpen		:= fbJaw.xRetracted;

IF fbJaw.xAlarm THEN
	M_RaiseAlarm(eNew := ALM_STK_JAW_TIMEOUT);
END_IF


// -------------------------------------------------------------
// 3. POPRAWNOSC POZYCJI
// -------------------------------------------------------------
//
// Pozycje wpisuje czlowiek, wiec sprawdzamy je zanim wozek
// ruszy. Musza tworzyc ciag - rosnacy albo malejacy.

IF NOT M_PositionsValid() THEN
	M_HaltDrive();
	M_RaiseAlarm(eNew := ALM_STK_POS_INVALID);
END_IF


// -------------------------------------------------------------
// 4. BLAD FALOWNIKA
// -------------------------------------------------------------

IF pDrive <> 0 THEN
	IF pDrive^.xFault OR pDrive^.xCommError THEN
		M_RaiseAlarm(eNew := ALM_STK_DRIVE_FAULT);
	END_IF
END_IF


// -------------------------------------------------------------
// 5. ZEZWOLENIE I TRYBY
// -------------------------------------------------------------

IF NOT xSafetyOK THEN
	M_HaltDrive();
	tonMoveWd(IN := FALSE);
	M_ApplyDrive();
	RETURN;
END_IF

IF xAlarm THEN
	M_HaltDrive();
	tonMoveWd(IN := FALSE);
	M_ApplyDrive();
	RETURN;
END_IF

IF eMode = MODE_MANUAL THEN
	M_ManualCycle();
	M_ApplyDrive();
	RETURN;
END_IF


// -------------------------------------------------------------
// 6. DOJAZD DO POZYCJI
// -------------------------------------------------------------

IF nTargetSel = 0 THEN
	M_HaltDrive();
	tonMoveWd(IN := FALSE);
	M_ApplyDrive();
	RETURN;
END_IF


IF ABS(diError) <= pP^.Cfg.diWindow THEN

	M_HaltDrive();
	tonMoveWd(IN := FALSE);

	// Krotkie uspokojenie, zanim stacja ruszy szczekami
	tonSettle(IN := TRUE, PT := pP^.Cfg.tSettle);
	xInPosition := tonSettle.Q;

	M_ApplyDrive();
	RETURN;

END_IF


xInPosition := FALSE;
tonSettle(IN := FALSE);


// Predkosc: pelna do strefy dojazdowej, potem dojazdowa
IF ABS(diError) > pP^.Cfg.diSlowZone THEN
	lrFreqReq := pP^.Cfg.lrFreqFast;
ELSE
	lrFreqReq := pP^.Cfg.lrFreqSlow;
END_IF


// Kierunek: znak bledu plus informacja, w ktora strone rosnie
// wskazanie enkodera
xRunReq := TRUE;

IF diError > 0 THEN
	xRevReq := NOT pP^.Cfg.xIncreaseIsForward;
ELSE
	xRevReq := pP^.Cfg.xIncreaseIsForward;
END_IF


// Watchdog dojazdu
tonMoveWd(IN := TRUE, PT := pP^.Cfg.tMoveWatchdog);

IF tonMoveWd.Q THEN
	M_HaltDrive();
	M_RaiseAlarm(eNew := ALM_STK_MOVE_TIMEOUT);
END_IF


M_ApplyDrive();

METHOD PUBLIC M_Config
// Wolac raz, przy starcie.
VAR_INPUT
	pPersist	: POINTER TO ST_StackPersist;
	pDrv		: POINTER TO FB_NordSK550PP;
	nJawId		: INT;
	pJawPersist	: POINTER TO ST_CylPersist;
END_VAR
pP		:= pPersist;
pDrive	:= pDrv;

fbJaw.M_Config(nId := nJawId, pPersist := pJawPersist);
END_METHOD

METHOD PUBLIC M_MoveTo : BOOL
// Zadanie pozycji. Zwraca TRUE, gdy wozek juz w niej stoi.
//   1 dol, 2 srodek, 3 gora
VAR_INPUT
	nSel	: INT;
END_VAR
M_MoveTo := FALSE;

IF pP = 0 THEN
	RETURN;
END_IF

IF nSel <> nTargetSel THEN
	nTargetSel := nSel;
	tonMoveWd(IN := FALSE);
	tonSettle(IN := FALSE);
	xInPosition := FALSE;
END_IF

CASE nSel OF
	1: diTarget := pP^.Cfg.diPosBottom;
	2: diTarget := pP^.Cfg.diPosMiddle;
	3: diTarget := pP^.Cfg.diPosTop;
ELSE
	nTargetSel := 0;
	RETURN;
END_CASE

M_MoveTo := xInPosition;
END_METHOD

METHOD PUBLIC M_Park
// Zdjecie zadania pozycji - wozek stoi tam, gdzie jest.
nTargetSel	:= 0;
xInPosition	:= FALSE;
tonMoveWd(IN := FALSE);
tonSettle(IN := FALSE);
END_METHOD

METHOD PUBLIC M_JawsClose : BOOL
// Zamkniecie szczek - wsuniecie ich w deski palety.
// Zwraca TRUE po potwierdzeniu.
fbJaw.M_Extend();
M_JawsClose := fbJaw.xExtended;
END_METHOD

METHOD PUBLIC M_JawsOpen : BOOL
fbJaw.M_Retract();
M_JawsOpen := fbJaw.xRetracted;
END_METHOD

METHOD PUBLIC M_ManJog
// Jazda reczna wozkiem oraz reczne szczeki.
VAR_INPUT
	xUp			: BOOL;
	xDown		: BOOL;
	xJawClose	: BOOL;
	xJawOpen	: BOOL;
END_VAR
xManUp		:= xUp;
xManDown	:= xDown;

fbJaw.M_ManJog(xExt := xJawClose, xRet := xJawOpen);
END_METHOD

METHOD PUBLIC M_Reset : BOOL
fbJaw.M_Reset();

IF pDrive <> 0 THEN
	pDrive^.M_Reset();
END_IF

eAlarm	:= ALM_STK_NONE;
xAlarm	:= FALSE;

tonMoveWd(IN := FALSE);
tonSettle(IN := FALSE);

nTargetSel	:= 0;
xInPosition	:= FALSE;
M_Reset		:= TRUE;
END_METHOD

METHOD PROTECTED M_PositionsValid : BOOL
// Dol, srodek i gora musza lezec po kolei. Odleglosc miedzy
// nimi to wysokosc palety, wiec pomylka w kolejnosci wyslalaby
// wozek w przeciwna strone niz trzeba.
VAR
	a	: DINT;
	b	: DINT;
	c	: DINT;
END_VAR
M_PositionsValid := FALSE;

a := pP^.Cfg.diPosBottom;
b := pP^.Cfg.diPosMiddle;
c := pP^.Cfg.diPosTop;

IF (a < b) AND (b < c) THEN
	M_PositionsValid := TRUE;
	RETURN;
END_IF

IF (a > b) AND (b > c) THEN
	M_PositionsValid := TRUE;
END_IF
END_METHOD

METHOD PROTECTED M_ManualCycle
// Jazda reczna bez pozycjonowania. Progi pozycji sa nadal
// pokazywane, ale nic nie zatrzymuje wozka za operatora.
nTargetSel	:= 0;
xInPosition	:= FALSE;
tonMoveWd(IN := FALSE);

IF xManUp AND NOT xManDown THEN
	xRunReq		:= TRUE;
	xRevReq		:= NOT pP^.Cfg.xIncreaseIsForward;
	lrFreqReq	:= pP^.Cfg.lrFreqManual;
	RETURN;
END_IF

IF xManDown AND NOT xManUp THEN
	xRunReq		:= TRUE;
	xRevReq		:= pP^.Cfg.xIncreaseIsForward;
	lrFreqReq	:= pP^.Cfg.lrFreqManual;
	RETURN;
END_IF

M_HaltDrive();
END_METHOD

METHOD PROTECTED M_HaltDrive
xRunReq		:= FALSE;
lrFreqReq	:= 0.0;
xMoving		:= FALSE;
END_METHOD

METHOD PROTECTED M_ApplyDrive
// Metody falownika wolamy na zboczu - blok napedu przy
// blokadzie sam kasuje zadanie ruchu i nie wolno mu go
// wracac samoczynnie.
xMoving := xRunReq;

IF pDrive = 0 THEN
	RETURN;
END_IF


IF xRunReq AND NOT xRunOld THEN
	pDrive^.M_Start(lrFreq := lrFreqReq, xReverse := xRevReq);
	xRevOld		:= xRevReq;
	lrFreqOld	:= lrFreqReq;
	xRunOld		:= xRunReq;
	RETURN;
END_IF

IF NOT xRunReq AND xRunOld THEN
	pDrive^.M_Stop();
	xRunOld := xRunReq;
	RETURN;
END_IF

IF NOT xRunReq THEN
	xRunOld := xRunReq;
	RETURN;
END_IF


IF xRevReq <> xRevOld THEN
	pDrive^.M_Start(lrFreq := lrFreqReq, xReverse := xRevReq);
	xRevOld		:= xRevReq;
	lrFreqOld	:= lrFreqReq;
	RETURN;
END_IF

IF lrFreqReq <> lrFreqOld THEN
	pDrive^.M_SetFrequency(lrFreq := lrFreqReq);
	lrFreqOld := lrFreqReq;
END_IF
END_METHOD

METHOD PROTECTED M_RaiseAlarm
VAR_INPUT
	eNew	: E_StackAlarm;
END_VAR
IF eNew = ALM_STK_NONE THEN
	RETURN;
END_IF

IF eAlarm = ALM_STK_NONE THEN
	eAlarm := eNew;
END_IF

xAlarm := TRUE;
END_METHOD

END_FUNCTION_BLOCK

// ---- POUs/POUs/FB/FB_Cylinder.TcPOU
FUNCTION_BLOCK FB_Cylinder
// =============================================================
// SILOWNIK PNEUMATYCZNY
// =============================================================
//
// Jeden blok na wszystkie silowniki maszyny - blokade stacji 5,
// szczeki, silowniki rozrywajace, dociski stacji 4, podnoszenie
// rolek na stacjach 8 i 10. Roznice siedza w nastawach, nie
// w kodzie.
//
// -------------------------------------------------------------
// ZAWORY
// -------------------------------------------------------------
// Blok wystawia dwie cewki: xCoilExtend i xCoilRetract. Stacja
// przepisuje je na swoje wyjscia. Sposob ich uzycia zalezy od
// typu zaworu (E_CylValve) - monostabilny uzywa tylko pierwszej,
// 3-polozeniowy w spoczynku ma zdjete obie.
//
// -------------------------------------------------------------
// SPRZEZENIE
// -------------------------------------------------------------
// Trzy warianty: brak, krancowki, przetwornik IO-Link o wartosci
// bezwzglednej. Przy przetworniku polozenia koncowe to PROGI
// nastawiane przez operatora, liczone wzgledem punktu bazowania.
//
// Obserwacje polozenia mozna wylaczyc OSOBNO dla kazdego
// kierunku i zastapic czasowka - tryb pracy z uszkodzonym
// czujnikiem. Tak samo watchdog: silownik bez krancowki na
// jednym koncu nie ma jak potwierdzic dojazdu, wiec watchdog
// w tym kierunku musi dac sie wylaczyc.
//
// -------------------------------------------------------------
// PRZEKROCZENIE PROGU
// -------------------------------------------------------------
// xOverLimit NIE JEST ALARMEM SILOWNIKA. To wynik testu:
// silownik wysunal sie dalej, niz moglby z cala paleta, czyli
// deska pekla albo odpadla. Decyzje podejmuje stacja.
VAR_INPUT

	eMode			: E_MachineMode;
	xSafetyOK		: BOOL;

	// Krancowki - logika dodatnia (TRUE = czujnik zadziala)
	xSwExtRaw		: BOOL;
	xSwRetRaw		: BOOL;

	// Surowe wskazanie przetwornika IO-Link
	diPosRaw		: DINT;

	// Sprzezenie z zewnatrz (CYLFB_EXTERNAL). Stacja 4 steruje
	// grupami silownikow jednym zaworem, a mierzy kazdy osobno -
	// agreguje wskazania monitorow i podaje wynik tutaj.
	xFbExtIn		: BOOL;
	xFbRetIn		: BOOL;

END_VAR
VAR_OUTPUT

	// Cewki zaworu - stacja przepisuje je na swoje wyjscia
	xCoilExtend		: BOOL;
	xCoilRetract	: BOOL;

	eState			: E_CylState;
	eAlarm			: E_CylAlarm;
	xAlarm			: BOOL;

	// Potwierdzone polozenia koncowe
	xExtended		: BOOL;
	xRetracted		: BOOL;
	xMoving			: BOOL;

	// Polozenie wzgledem punktu bazowania
	diPos			: DINT;

	// Przekroczenie progu = deska pekla / odpadla
	xOverLimit		: BOOL;

	// Nacisk utrzymany przez nastawiony czas (stacja 5)
	xHoldDone		: BOOL;

END_VAR
VAR

	nCylId			: INT;
	pP				: POINTER TO ST_CylPersist;

	// Zadanie: TRUE = wysuw
	xReqExtend		: BOOL;
	xCmdIssued		: BOOL;

	// Sprzezenie po odfiltrowaniu wylaczen
	xFbExtended		: BOOL;
	xFbRetracted	: BOOL;
	xFbConflict		: BOOL;

	tonDelay		: TON;
	tonWatchdog		: TON;
	tonSubst		: TON;
	tonSettle		: TON;
	tonHold			: TON;

	eModeOld		: E_MachineMode;

	xManExtend		: BOOL;
	xManRetract		: BOOL;

END_VAR

// =============================================================
// CYKL SILOWNIKA
// =============================================================


// -------------------------------------------------------------
// 1. KONFIGURACJA
// -------------------------------------------------------------

IF pP = 0 THEN
	M_Deenergize();
	eAlarm	:= ALM_CYL_NOT_CONFIGURED;
	xAlarm	:= TRUE;
	eState	:= CYL_ALARM;
	RETURN;
END_IF


// -------------------------------------------------------------
// 2. POLOZENIE I SPRZEZENIE
// -------------------------------------------------------------

M_ReadPosition();
M_EvalFeedback();

// Potwierdzone polozenia koncowe bierzemy ze STANU, nie wprost
// z czujnika. Dzieki temu dzialaja tak samo wtedy, gdy operator
// wylaczyl obserwacje czujnika i ruch potwierdza czasowka.
xExtended	:= (eState = CYL_EXTENDED);
xRetracted	:= (eState = CYL_RETRACTED);
xAlarm		:= (eAlarm <> ALM_CYL_NONE);


// -------------------------------------------------------------
// 3. NIEZGODNOSC KRANCOWEK
// -------------------------------------------------------------

tonSettle(IN := xFbConflict, PT := pP^.Cfg.tSettle);

IF tonSettle.Q THEN
	M_RaiseAlarm(eNew := ALM_CYL_BOTH_SWITCHES);
END_IF


// -------------------------------------------------------------
// 4. ZEZWOLENIE BEZPIECZENSTWA
// -------------------------------------------------------------
//
// Cewki zostaja tam, gdzie byly - zdjecie ich przy zaworze
// monostabilnym cofneloby silownik, a to przy zamknietych
// szczekach na palecie nie jest bezpieczne. Ruch stoi,
// watchdog jest wyzerowany i po powrocie zezwolenia liczy
// od poczatku.

IF NOT xSafetyOK THEN
	xMoving := FALSE;
	tonWatchdog(IN := FALSE);
	tonSubst(IN := FALSE);
	tonDelay(IN := FALSE);
	RETURN;
END_IF


// -------------------------------------------------------------
// 5. TRYB RECZNY
// -------------------------------------------------------------

IF eMode = MODE_MANUAL THEN
	eModeOld := eMode;
	M_ManualCycle();
	RETURN;
END_IF

IF eModeOld = MODE_MANUAL THEN
	// Po recznej nie wiemy, gdzie operator zostawil silownik
	eState := CYL_UNKNOWN;
END_IF

eModeOld := eMode;


// -------------------------------------------------------------
// 6. ALARM
// -------------------------------------------------------------

IF xAlarm THEN
	xMoving	:= FALSE;
	eState	:= CYL_ALARM;
	RETURN;
END_IF


// -------------------------------------------------------------
// 7. SEKWENCJA
// -------------------------------------------------------------

CASE eState OF

CYL_UNKNOWN:
	xMoving := FALSE;

	IF NOT xCmdIssued THEN
		// Bez komendy nie ruszamy - nie wiadomo, co stoi na drodze
		RETURN;
	END_IF

	M_BeginMove(xExt := xReqExtend);


CYL_RETRACTED:
	xMoving := FALSE;
	M_ApplyCoils(xExt := FALSE);

	IF xReqExtend THEN
		M_BeginMove(xExt := TRUE);
	END_IF


CYL_EXTENDING:
	xMoving := TRUE;
	M_MoveCycle(xExt := TRUE);


CYL_EXTENDED:
	xMoving := FALSE;
	M_ApplyCoils(xExt := TRUE);

	IF NOT xReqExtend THEN
		M_BeginMove(xExt := FALSE);
	END_IF


CYL_RETRACTING:
	xMoving := TRUE;
	M_MoveCycle(xExt := FALSE);


CYL_ALARM:
	xMoving := FALSE;


ELSE
	eState := CYL_UNKNOWN;

END_CASE


// Odswiezenie po zmianie stanu w tym cyklu
xExtended	:= (eState = CYL_EXTENDED);
xRetracted	:= (eState = CYL_RETRACTED);


// -------------------------------------------------------------
// 8. TEST TRZYMANIA NACISKU
// -------------------------------------------------------------
//
// Liczymy czas dopiero od momentu, w ktorym silownik przekroczyl
// zaprogramowana pozycje. Kazdy silownik ma wlasny licznik, bo
// wszystkie ida z inna predkoscia.

IF pP^.Cfg.eFeedback = CYLFB_ANALOG THEN
	tonHold(IN := (diPos >= pP^.Cfg.diPosHoldStart), PT := pP^.Cfg.tHold);
	xHoldDone := tonHold.Q;
ELSE
	tonHold(IN := FALSE);
	xHoldDone := FALSE;
END_IF

METHOD PUBLIC M_Config
VAR_INPUT
	nId			: INT;
	pPersist	: POINTER TO ST_CylPersist;
END_VAR
nCylId	:= nId;
pP		:= pPersist;
END_METHOD

METHOD PUBLIC M_Extend : BOOL
// Zadanie wysuwu. Zatrzaskiwane - obowiazuje az do M_Retract.
xReqExtend	:= TRUE;
xCmdIssued	:= TRUE;
M_Extend	:= TRUE;
END_METHOD

METHOD PUBLIC M_Retract : BOOL
xReqExtend	:= FALSE;
xCmdIssued	:= TRUE;
M_Retract	:= TRUE;
END_METHOD

METHOD PUBLIC M_ManJog
// Komendy trybu recznego. Dzialaja tylko w MODE_MANUAL.
VAR_INPUT
	xExt	: BOOL;
	xRet	: BOOL;
END_VAR
xManExtend	:= xExt;
xManRetract	:= xRet;
END_METHOD

METHOD PUBLIC M_Zero : BOOL
// Bazowanie przetwornika w BIEZACYM polozeniu.
//
// Stacja 4: wstawiamy palete, wysuwamy wszystkie silowniki
// i zerujemy - punkt bazowy jest na silowniku WYSUNIETYM.
// Stacja 5: zerujemy na silowniku WYCOFANYM, bez palety.
//
// Dozwolone tylko w trybie recznym.
M_Zero := FALSE;

IF pP = 0 THEN
	RETURN;
END_IF

IF eMode <> MODE_MANUAL THEN
	RETURN;
END_IF

IF pP^.Cfg.eFeedback <> CYLFB_ANALOG THEN
	RETURN;
END_IF

pP^.Mem.diZeroOffset	:= diPosRaw;
pP^.Mem.xZeroed			:= TRUE;

M_Zero := TRUE;
END_METHOD

METHOD PUBLIC M_Reset : BOOL
eAlarm	:= ALM_CYL_NONE;
xAlarm	:= FALSE;

tonWatchdog(IN := FALSE);
tonSubst(IN := FALSE);
tonDelay(IN := FALSE);
tonSettle(IN := FALSE);

eState	:= CYL_UNKNOWN;
M_Reset	:= TRUE;
END_METHOD

METHOD PROTECTED M_ReadPosition
// Przeliczenie wskazania surowego na polozenie wzgledem bazy.
// Znak dodatni zawsze w kierunku wysuwu.
IF pP^.Cfg.eFeedback <> CYLFB_ANALOG THEN
	diPos := 0;
	RETURN;
END_IF

IF pP^.Cfg.xInvertPos THEN
	diPos := pP^.Mem.diZeroOffset - diPosRaw;
	RETURN;
END_IF

diPos := diPosRaw - pP^.Mem.diZeroOffset;
END_METHOD

METHOD PROTECTED M_EvalFeedback
xOverLimit := FALSE;

CASE pP^.Cfg.eFeedback OF

CYLFB_SWITCHES:
	xFbExtended		:= xSwExtRaw;
	xFbRetracted	:= xSwRetRaw;
	xFbConflict		:= xSwExtRaw AND xSwRetRaw;

CYLFB_ANALOG:
	xFbExtended		:= (diPos >= pP^.Cfg.diPosExtended);
	xFbRetracted	:= (diPos <= pP^.Cfg.diPosRetracted);
	xFbConflict		:= FALSE;
	xOverLimit		:= (diPos > pP^.Cfg.diPosLimit);

CYLFB_EXTERNAL:
	xFbExtended		:= xFbExtIn;
	xFbRetracted	:= xFbRetIn;
	xFbConflict		:= xFbExtIn AND xFbRetIn;

ELSE
	// CYLFB_NONE - ruch wylacznie na czasowkach
	xFbExtended		:= FALSE;
	xFbRetracted	:= FALSE;
	xFbConflict		:= FALSE;

END_CASE
END_METHOD

METHOD PROTECTED M_BeginMove
VAR_INPUT
	xExt	: BOOL;
END_VAR
tonDelay(IN := FALSE);
tonWatchdog(IN := FALSE);
tonSubst(IN := FALSE);

IF xExt THEN
	eState := CYL_EXTENDING;
	RETURN;
END_IF

eState := CYL_RETRACTING;
END_METHOD

METHOD PROTECTED M_MoveCycle
// Jeden ruch: opoznienie -> wysterowanie zaworu ->
// potwierdzenie konca -> watchdog.
VAR_INPUT
	xExt		: BOOL;
END_VAR
VAR
	tDelay		: TIME;
	tSubst		: TIME;
	tWd			: TIME;
	xFbUsed		: BOOL;
	xFbReached	: BOOL;
	xWdEnabled	: BOOL;
	xDone		: BOOL;
END_VAR
// ---------------------------------------------------------
// Nastawy dla biezacego kierunku
// ---------------------------------------------------------

IF xExt THEN
	tDelay		:= pP^.Cfg.tExtendDelay;
	tSubst		:= pP^.Cfg.tExtendSubst;
	tWd			:= pP^.Cfg.tExtendWatchdog;
	xFbUsed		:= pP^.Cfg.xExtendFbEnabled;
	xWdEnabled	:= pP^.Cfg.xExtendWdEnabled;
	xFbReached	:= xFbExtended;
ELSE
	tDelay		:= pP^.Cfg.tRetractDelay;
	tSubst		:= pP^.Cfg.tRetractSubst;
	tWd			:= pP^.Cfg.tRetractWatchdog;
	xFbUsed		:= pP^.Cfg.xRetractFbEnabled;
	xWdEnabled	:= pP^.Cfg.xRetractWdEnabled;
	xFbReached	:= xFbRetracted;
END_IF


// ---------------------------------------------------------
// Opoznienie wysterowania zaworu
// ---------------------------------------------------------
//
// W tej fazie NIE ruszamy cewek - silownik zostaje tam,
// gdzie byl. Zdjecie cewki zaworu monostabilnego cofneloby
// go, a o to nam nie chodzi.

tonDelay(IN := TRUE, PT := tDelay);

IF NOT tonDelay.Q THEN
	RETURN;
END_IF


// ---------------------------------------------------------
// Wysterowanie zaworu
// ---------------------------------------------------------

M_ApplyCoils(xExt := xExt);


// ---------------------------------------------------------
// Potwierdzenie konca ruchu
// ---------------------------------------------------------
//
// Sprzezenie wylaczone przez operatora = uznajemy ruch za
// wykonany po uplywie czasowki zastepczej.

IF xFbUsed THEN
	tonSubst(IN := FALSE);
	xDone := xFbReached;
ELSE
	tonSubst(IN := TRUE, PT := tSubst);
	xDone := tonSubst.Q;
END_IF


IF xDone THEN
	tonWatchdog(IN := FALSE);
	tonSubst(IN := FALSE);
	tonDelay(IN := FALSE);

	IF xExt THEN
		eState := CYL_EXTENDED;
	ELSE
		eState := CYL_RETRACTED;
	END_IF

	RETURN;
END_IF


// ---------------------------------------------------------
// Watchdog
// ---------------------------------------------------------
//
// Wylaczalny osobno dla kierunku bez krancowki.

tonWatchdog(IN := xWdEnabled, PT := tWd);

IF NOT tonWatchdog.Q THEN
	RETURN;
END_IF

IF xExt THEN
	M_RaiseAlarm(eNew := ALM_CYL_EXTEND_TIMEOUT);
	RETURN;
END_IF

M_RaiseAlarm(eNew := ALM_CYL_RETRACT_TIMEOUT);
END_METHOD

METHOD PROTECTED M_ApplyCoils
VAR_INPUT
	xExt	: BOOL;
END_VAR
CASE pP^.Cfg.eValve OF

CYLV_SINGLE:
	// Jedna cewka, powrot sprezyna
	xCoilExtend		:= xExt;
	xCoilRetract	:= FALSE;

CYLV_3POS_OFF_RET:
	// Cofniecie realizuje zdjecie cewek
	xCoilExtend		:= xExt;
	xCoilRetract	:= FALSE;

ELSE
	// CYLV_DOUBLE i CYLV_3POS_MID - cewki wykluczajace sie
	xCoilExtend		:= xExt;
	xCoilRetract	:= NOT xExt;

END_CASE
END_METHOD

METHOD PROTECTED M_Deenergize
// Zdjecie obu cewek. Przy zaworze 3-polozeniowym to jest
// polozenie spoczynkowe, przy monostabilnym powrot sprezyna.
xCoilExtend		:= FALSE;
xCoilRetract	:= FALSE;
END_METHOD

METHOD PROTECTED M_RaiseAlarm
// Pierwszy alarm zostaje - operator ma widziec przyczyne.
VAR_INPUT
	eNew	: E_CylAlarm;
END_VAR
IF eNew = ALM_CYL_NONE THEN
	RETURN;
END_IF

IF eAlarm = ALM_CYL_NONE THEN
	eAlarm := eNew;
END_IF

xAlarm	:= TRUE;
eState	:= CYL_ALARM;
xMoving	:= FALSE;
END_METHOD

METHOD PROTECTED M_ManualCycle
// Praca reczna: sterowanie cewkami wprost, bez watchdogow
// i bez czasowek. Sluzy takze do bazowania przetwornikow.
eState := CYL_MANUAL;

tonWatchdog(IN := FALSE);
tonSubst(IN := FALSE);
tonDelay(IN := FALSE);

IF xManExtend AND NOT xManRetract THEN
	M_ApplyCoils(xExt := TRUE);
	xMoving := TRUE;
	RETURN;
END_IF

IF xManRetract AND NOT xManExtend THEN
	M_ApplyCoils(xExt := FALSE);
	xMoving := TRUE;
	RETURN;
END_IF

xMoving := FALSE;
END_METHOD

END_FUNCTION_BLOCK

// ---- POUs/POUs/FB/FB_Station03_Destack.TcPOU
FUNCTION_BLOCK FB_Station03_Destack EXTENDS FB_RollerConveyor
// =============================================================
// STACJA 3 - DESZTAPLARKA
// =============================================================
//
// Rozdziela stos na pojedyncze palety. Wozek ze szczekami chwyta
// pod DRUGA palete od dolu i unosi caly stos - najnizsza paleta
// zostaje na transporterze i moze wyjechac.
//
// -------------------------------------------------------------
// CYKL
// -------------------------------------------------------------
//   w trakcie wjazdu   szczeki otwarte, wozek jedzie na SRODEK
//   po potwierdzeniu   zapamietanie, ze stos dojechal
//   chwyt              szczeki zamykaja sie pod druga paleta
//   uniesienie         wozek na GORE, dolna paleta wolna
//   wydanie            paleta wyjezdza na stacje 4
//   odlozenie          wozek na DOL, szczeki otwarte
//   i od nowa, az stos sie skonczy
//
// -------------------------------------------------------------
// OSTATNIA PALETA
// -------------------------------------------------------------
// Gdy na transporterze zostaje JEDNA paleta, nie ma juz czego
// chwytac - nie ma drugiej palety od dolu. Ostatnia sztuka
// wyjezdza wprost z transportera, bez unoszenia.
//
// -------------------------------------------------------------
// LICZBA PALET
// -------------------------------------------------------------
// Na razie stala, z Cfg.nStackSize. Czujnik wykrywajacy, ze stos
// sie skonczyl, dojdzie pozniej - wtedy licznik bedzie tylko
// wartoscia oczekiwana, a prawde powie czujnik.
VAR_INPUT

	// Enkoder absolutny wozka
	diLiftPosRaw	: DINT;

	// Krancowki szczek
	xJawClosedSw	: BOOL;
	xJawOpenSw		: BOOL;

END_VAR
VAR_OUTPUT

	// Cewki szczek - stacja przepisuje je na swoje wyjscia
	xJawCoilClose	: BOOL;
	xJawCoilOpen	: BOOL;

	nStep			: INT;

	// Ile palet zostalo do wydania z biezacego stosu
	nRemaining		: INT;

	diLiftPos		: DINT;
	nLiftTarget		: INT;
	xLiftInPos		: BOOL;

	eLiftAlarm		: E_StackAlarm;

END_VAR
VAR

	pSt		: POINTER TO ST_StackPersist;
	fbLift	: FB_StackLift;

	nNextId	: UDINT;

END_VAR
VAR CONSTANT

	ST3_IDLE		: INT := 0;
	ST3_PREPOS		: INT := 10;
	ST3_GRIP		: INT := 20;
	ST3_LIFT		: INT := 30;
	ST3_HANDOVER	: INT := 40;
	ST3_WAIT_CLEAR	: INT := 50;
	ST3_LOWER		: INT := 60;
	ST3_OPEN		: INT := 70;
	ST3_LAST		: INT := 80;
	ST3_EMPTYSTACK	: INT := 90;

END_VAR

// =============================================================
// CYKL STACJI 3
// =============================================================


// 1. Wozek ze szczekami
M_CallLift();


// 2. Warstwa transportu
SUPER^();


// 3. Sekwencja desztaplowania.
//    Chodzi w KAZDYM stanie wezla, nie tylko w NODE_BUSY:
//    odkladanie stosu i chwyt nastepnej palety odbywaja sie
//    wtedy, gdy wezel jest juz pusty po wydaniu poprzedniej.
M_DestackCycle();


// 4. Diagnostyka
M_MapStatus();

METHOD PUBLIC M_ConfigStation
// Wolac raz, przy starcie, PO M_Config klasy bazowej.
VAR_INPUT
	pStPersist	: POINTER TO ST_StackPersist;

	// Falownik 1 - krzywka desztaplarki
	pLiftDrive	: POINTER TO FB_NordSK550PP;

	// Rekord silownika szczek
	nJawId		: INT;
	pJawPersist	: POINTER TO ST_CylPersist;
END_VAR
pSt := pStPersist;

fbLift.M_Config(
	pPersist	:= pStPersist,
	pDrv		:= pLiftDrive,
	nJawId		:= nJawId,
	pJawPersist	:= pJawPersist
);
END_METHOD

METHOD PROTECTED M_CallLift
fbLift(
	eMode			:= eMode,
	xSafetyOK		:= xSafetyOK,
	diPosRaw		:= diLiftPosRaw,
	xJawClosedSw	:= xJawClosedSw,
	xJawOpenSw		:= xJawOpenSw
);

xJawCoilClose	:= fbLift.xJawCoilClose;
xJawCoilOpen	:= fbLift.xJawCoilOpen;

IF fbLift.xAlarm THEN
	M_RaiseAlarm(eNew := ALM_OPERATION_FAILED);
END_IF
END_METHOD

METHOD PROTECTED M_MapStatus
diLiftPos	:= fbLift.diPos;
nLiftTarget	:= fbLift.nTargetSel;
xLiftInPos	:= fbLift.xInPosition;
eLiftAlarm	:= fbLift.eAlarm;

IF pSt <> 0 THEN
	nRemaining := pSt^.Mem.nRemaining;
END_IF
END_METHOD

METHOD PUBLIC M_StackArrived : BOOL
// Stos dojechal do pozycji i zostal potwierdzony czujnikami.
//
// Liczbe palet zapisujemy W PAMIECI NIEULOTNEJ - po zaniku
// zasilania maszyna musi wiedziec, ile sztuk zostalo jeszcze
// w stosie stojacym na stacji.
M_StackArrived := FALSE;

IF pSt = 0 THEN
	RETURN;
END_IF

IF pSt^.Mem.xStackArrived THEN
	RETURN;
END_IF

pSt^.Mem.xStackArrived	:= TRUE;
pSt^.Mem.nRemaining		:= pSt^.Cfg.nStackSize;
xPersistDirty			:= TRUE;

M_StackArrived := TRUE;
END_METHOD

METHOD PROTECTED M_OperationRequired : BOOL
// Stos musi sie zatrzymac i zostac rozdzielony. Pojedyncza
// paleta wydana przez desztaplarke jest juz obsluzona -
// M_InjectLoad ustawia jej xOperationDone.
M_OperationRequired := TRUE;

IF pP = 0 THEN
	RETURN;
END_IF

IF NOT pP^.Cfg.xStationEnabled THEN
	M_OperationRequired := FALSE;
	RETURN;
END_IF

M_OperationRequired := NOT pP^.Mem.xOperationDone;
END_METHOD

METHOD PROTECTED M_OperationCycle : BOOL
// Wezel czeka, az desztaplarka odseparuje pierwsza palete.
// Wlasciwa sekwencja siedzi w M_DestackCycle, bo musi dzialac
// takze wtedy, gdy wezel jest pusty.
M_OperationCycle := FALSE;

IF pP = 0 THEN
	RETURN;
END_IF

M_OperationCycle := pP^.Mem.xOperationDone;
END_METHOD

METHOD PROTECTED M_TravelCycle
// W trakcie wjazdu stosu wozek ma byc otwarty i stac na
// pozycji chwytu - zeby po potwierdzeniu czujnikami od razu
// mozna bylo zamknac szczeki.
IF nStep <> ST3_IDLE THEN
	RETURN;
END_IF

fbLift.M_JawsOpen();
fbLift.M_MoveTo(nSel := 2);
END_METHOD

METHOD PROTECTED M_DestackCycle
// Sekwencja desztaplowania.
IF pSt = 0 THEN
	RETURN;
END_IF

IF pP = 0 THEN
	RETURN;
END_IF

IF NOT xSafetyOK THEN
	RETURN;
END_IF

IF xAlarm THEN
	RETURN;
END_IF

IF eMode <> MODE_AUTO THEN
	RETURN;
END_IF

// Stacja wylaczona przez operatora - stos przejezdza w calosci,
// bez rozdzielania. Uzywane przy uruchomieniu transportu.
IF NOT pP^.Cfg.xStationEnabled THEN
	nStep := ST3_IDLE;
	RETURN;
END_IF


CASE nStep OF

ST3_IDLE:
	// Czekamy, az stos zatrzyma sie na czujnikach
	IF NOT pP^.Mem.xLoadPresent THEN
		RETURN;
	END_IF

	IF (eState <> NODE_BUSY) AND (eState <> NODE_OCCUPIED) THEN
		RETURN;
	END_IF

	M_StackArrived();

	IF pSt^.Mem.nRemaining <= 1 THEN
		nStep := ST3_LAST;
		RETURN;
	END_IF

	nStep := ST3_PREPOS;


ST3_PREPOS:
	// Szczeki otwarte, wozek pod druga palete od dolu
	fbLift.M_JawsOpen();

	IF NOT fbLift.xJawsOpen THEN
		RETURN;
	END_IF

	IF fbLift.M_MoveTo(nSel := 2) THEN
		nStep := ST3_GRIP;
	END_IF


ST3_GRIP:
	// Szczeki wchodza w deski drugiej palety od dolu
	IF fbLift.M_JawsClose() THEN
		pSt^.Mem.xJawsLoaded	:= TRUE;
		xPersistDirty			:= TRUE;
		nStep					:= ST3_LIFT;
	END_IF


ST3_LIFT:
	// Uniesienie stosu - najnizsza paleta zostaje na transporterze
	IF fbLift.M_MoveTo(nSel := 3) THEN
		nStep := ST3_HANDOVER;
	END_IF


ST3_HANDOVER:
	// Odseparowana paleta staje sie ladunkiem wezla i moze jechac
	nNextId := pP^.Mem.nLoadId;
	M_InjectLoad(xNok := FALSE, nLoadId := nNextId, xOpDone := TRUE);
	nStep := ST3_WAIT_CLEAR;


ST3_WAIT_CLEAR:
	// Czekamy, az paleta zjedzie ze stacji
	IF pP^.Mem.xLoadPresent THEN
		RETURN;
	END_IF

	pSt^.Mem.nRemaining	:= pSt^.Mem.nRemaining - 1;
	xPersistDirty		:= TRUE;

	IF pSt^.Mem.nRemaining <= 0 THEN
		nStep := ST3_EMPTYSTACK;
		RETURN;
	END_IF

	nStep := ST3_LOWER;


ST3_LOWER:
	// Odlozenie stosu na transporter
	IF fbLift.M_MoveTo(nSel := 1) THEN
		nStep := ST3_OPEN;
	END_IF


ST3_OPEN:
	IF fbLift.M_JawsOpen() THEN
		pSt^.Mem.xJawsLoaded	:= FALSE;
		xPersistDirty			:= TRUE;

		// Ostatnia paleta nie ma nad soba drugiej - wyjezdza
		// wprost z transportera, bez unoszenia
		IF pSt^.Mem.nRemaining <= 1 THEN
			nStep := ST3_LAST;
			RETURN;
		END_IF

		nStep := ST3_PREPOS;
	END_IF


ST3_LAST:
	// Jedna paleta na transporterze - wydajemy ja bez chwytania
	fbLift.M_JawsOpen();
	fbLift.M_MoveTo(nSel := 2);

	nNextId := pP^.Mem.nLoadId;
	M_InjectLoad(xNok := FALSE, nLoadId := nNextId, xOpDone := TRUE);

	nStep := ST3_WAIT_CLEAR;


ST3_EMPTYSTACK:
	// Stos wydany w calosci - stacja gotowa na nastepny
	pSt^.Mem.xStackArrived	:= FALSE;
	pSt^.Mem.nRemaining		:= 0;
	pSt^.Mem.xJawsLoaded	:= FALSE;
	xPersistDirty			:= TRUE;

	fbLift.M_JawsOpen();
	fbLift.M_MoveTo(nSel := 2);

	nStep := ST3_IDLE;


ELSE
	nStep := ST3_IDLE;

END_CASE
END_METHOD

METHOD PROTECTED M_SensorCheckAllowed : BOOL
// Porownanie pamieci z czujnikami ma sens tylko wtedy, gdy to,
// co lezy na transporterze, jest ladunkiem wezla.
//
// W trakcie desztaplowania tak nie jest: stos wisi na szczekach
// albo wlasnie schodzi na transporter, a pamiec wezla mowi
// "pusto". Bez tego wyjatku maszyna zglaszalaby nieistniejacy
// blad przy kazdej palecie.
M_SensorCheckAllowed := (nStep = ST3_IDLE) OR (nStep = ST3_WAIT_CLEAR);
END_METHOD

METHOD PUBLIC M_Reset : BOOL
// Reset NIE kasuje licznika palet w stosie - stos fizycznie
// lezy na stacji i maszyna ma o nim pamietac. Do wyzerowania
// stanu sluzy M_ServiceClearStack.
fbLift.M_Reset();

M_Reset := SUPER^.M_Reset();
END_METHOD

METHOD PUBLIC M_ServiceClearStack : BOOL
// Serwis zabral stos recznie i potwierdza, ze stacja jest pusta.
M_ServiceClearStack := FALSE;

IF pSt = 0 THEN
	RETURN;
END_IF

pSt^.Mem.xStackArrived	:= FALSE;
pSt^.Mem.nRemaining		:= 0;
pSt^.Mem.xJawsLoaded	:= FALSE;
xPersistDirty			:= TRUE;

nStep := ST3_IDLE;

M_ServiceClearStack := M_ServiceSetEmpty();
END_METHOD

METHOD PUBLIC M_ManLift
VAR_INPUT
	xUp			: BOOL;
	xDown		: BOOL;
	xJawClose	: BOOL;
	xJawOpen	: BOOL;
END_VAR
fbLift.M_ManJog(
	xUp			:= xUp,
	xDown		:= xDown,
	xJawClose	:= xJawClose,
	xJawOpen	:= xJawOpen
);
END_METHOD

END_FUNCTION_BLOCK

// ---- POUs/POUs/FB/FB_RollerConveyor.TcPOU
FUNCTION_BLOCK FB_RollerConveyor EXTENDS FB_TransportNodeBase
// =============================================================
// TRANSPORTER ROLKOWY
// =============================================================
//
// Standardowy wezel maszyny: naped NORDAC PRO SK 550P plus dwa
// czujniki optyczne na koncu transportera.
//
// -------------------------------------------------------------
// CZUJNIKI
// -------------------------------------------------------------
// Logika ODWROCONA: sygnal 1 = wolne, sygnal 0 = cos widac.
// Obecnosc palety w pozycji koncowej to ZERO Z OBU czujnikow -
// sa ustawione geometrycznie tak, ze jeden widzi pierwsza,
// a drugi ostatnia kostke palety.
//
// W trakcie przejazdu kostki palety "migaja" pierwszym
// czujnikiem. Nie ma to znaczenia, bo pozycje uznajemy dopiero
// po zgodnym zeru z obu czujnikow.
//
// Kazdy czujnik operator moze wylaczyc z HMI (uszkodzony).
// Wylaczenie obu przelacza wezel na przejazd czasowkowy.
//
// -------------------------------------------------------------
// NAPED
// -------------------------------------------------------------
// FB nie wola metod napedu co cykl, tylko na zboczu zadania.
// FB_NordSK550PP przy blokadzie (blad, STO, komunikacja) sam
// kasuje zadanie ruchu - i naped NIE MOZE ruszyc sam po
// ustapieniu przyczyny. Wolanie M_Start co cykl zepsuloby
// to zabezpieczenie.
VAR_INPUT

	// Surowe sygnaly czujnikow, logika odwrocona
	xSens1Raw		: BOOL := TRUE;
	xSens2Raw		: BOOL := TRUE;

END_VAR
VAR_OUTPUT

	// Stan czujnikow po odwroceniu logiki i po uwzglednieniu
	// wylaczen - do podgladu na HMI
	xSens1Detect	: BOOL;
	xSens2Detect	: BOOL;

END_VAR
VAR

	pDrive			: POINTER TO FB_NordSK550PP;

	xRunOld			: BOOL;
	xRevOld			: BOOL;
	xRevOut			: BOOL;
	lrFreqOld		: LREAL;

END_VAR

// =============================================================
// CYKL TRANSPORTERA ROLKOWEGO
// =============================================================


// 1. Czujniki -> szew klasy bazowej
M_ReadSensors();


// 2. Stan napedu -> szew klasy bazowej
M_ReadDrive();


// 3. Wspolna logika wezla
SUPER^();


// 4. Zadanie klasy bazowej -> naped
M_ApplyDrive();

METHOD PUBLIC M_ConfigDrive
// Podpiecie falownika. Wolac raz, przy starcie.
VAR_INPUT
	pDrv	: POINTER TO FB_NordSK550PP;
END_VAR
pDrive := pDrv;
END_METHOD

METHOD PROTECTED M_ReadSensors
// Odwrocenie logiki i uwzglednienie wylaczen serwisowych.
VAR
	xS1	: BOOL;
	xS2	: BOOL;
END_VAR
IF pP = 0 THEN
	xSensUsable		:= FALSE;
	xSensLoadAtStop	:= FALSE;
	xSensLoadNone	:= FALSE;
	xSensConflict	:= FALSE;
	xSens1Detect	:= FALSE;
	xSens2Detect	:= FALSE;
	RETURN;
END_IF


// Polaryzacja czujnikow z nastaw - maszyna docelowa pracuje
// w logice odwroconej, wersja testowa wprost
IF pP^.Cfg.xSensorsInverted THEN
	xS1 := NOT xSens1Raw;
	xS2 := NOT xSens2Raw;
ELSE
	xS1 := xSens1Raw;
	xS2 := xSens2Raw;
END_IF

xSens1Detect := xS1 AND pP^.Cfg.xSensor1Enabled;
xSens2Detect := xS2 AND pP^.Cfg.xSensor2Enabled;


// --- oba czujniki sprawne ---
IF pP^.Cfg.xSensor1Enabled AND pP^.Cfg.xSensor2Enabled THEN
	xSensUsable		:= TRUE;
	xSensLoadAtStop	:= xS1 AND xS2;
	xSensLoadNone	:= NOT xS1 AND NOT xS2;
	xSensConflict	:= xS1 XOR xS2;
	RETURN;
END_IF


// --- pracuje tylko czujnik 1 ---
IF pP^.Cfg.xSensor1Enabled THEN
	xSensUsable		:= TRUE;
	xSensLoadAtStop	:= xS1;
	xSensLoadNone	:= NOT xS1;
	xSensConflict	:= FALSE;
	RETURN;
END_IF


// --- pracuje tylko czujnik 2 ---
IF pP^.Cfg.xSensor2Enabled THEN
	xSensUsable		:= TRUE;
	xSensLoadAtStop	:= xS2;
	xSensLoadNone	:= NOT xS2;
	xSensConflict	:= FALSE;
	RETURN;
END_IF


// --- oba wylaczone: przejazd na czasowke ---
xSensUsable		:= FALSE;
xSensLoadAtStop	:= FALSE;
xSensLoadNone	:= FALSE;
xSensConflict	:= FALSE;
END_METHOD

METHOD PROTECTED M_ReadDrive
IF pDrive = 0 THEN
	xDrvReady := FALSE;
	xDrvFault := FALSE;
	RETURN;
END_IF

xDrvFault := pDrive^.xFault OR pDrive^.xCommError;
xDrvReady := NOT pDrive^.xError;
END_METHOD

METHOD PROTECTED M_ApplyDrive
// Przepisanie zadania klasy bazowej na metody falownika.
// Wylacznie na zboczach - patrz komentarz w naglowku FB.
IF pDrive = 0 THEN
	RETURN;
END_IF

IF pP = 0 THEN
	RETURN;
END_IF


// Trwale odwrocenie kierunku dla zle podlaczonych silnikow
xRevOut := xDrvRev XOR pP^.Cfg.xInvertDirection;


// --- start ---
IF xDrvRun AND NOT xRunOld THEN
	pDrive^.M_Start(lrFreq := lrDrvFreq, xReverse := xRevOut);
	xRevOld		:= xRevOut;
	lrFreqOld	:= lrDrvFreq;
	xRunOld		:= xDrvRun;
	RETURN;
END_IF


// --- stop ---
IF NOT xDrvRun AND xRunOld THEN
	pDrive^.M_Stop();
	xRunOld := xDrvRun;
	RETURN;
END_IF


IF NOT xDrvRun THEN
	xRunOld := xDrvRun;
	RETURN;
END_IF


// --- zmiana kierunku w ruchu (tylko tryb reczny) ---
IF xRevOut <> xRevOld THEN
	pDrive^.M_Start(lrFreq := lrDrvFreq, xReverse := xRevOut);
	xRevOld		:= xRevOut;
	lrFreqOld	:= lrDrvFreq;
	RETURN;
END_IF


// --- zmiana zadanej czestotliwosci ---
IF lrDrvFreq <> lrFreqOld THEN
	pDrive^.M_SetFrequency(lrFreq := lrDrvFreq);
	lrFreqOld := lrDrvFreq;
END_IF
END_METHOD

METHOD PUBLIC M_Reset : BOOL
// Reset wezla plus kasowanie bledu falownika.
IF pDrive <> 0 THEN
	pDrive^.M_Reset();
END_IF

M_Reset := SUPER^.M_Reset();
END_METHOD

END_FUNCTION_BLOCK

// ---- POUs/POUs/FB/FB_TransportNodeBase.TcPOU
FUNCTION_BLOCK FB_TransportNodeBase
// =============================================================
// WEZEL TRANSPORTU - KLASA BAZOWA
// =============================================================
//
// Wspolne dla wszystkich 16 stacji: pamiec obecnosci w
// zmiennych nieulotnych, weryfikacja pamieci wzgledem
// czujnikow, watchdogi przejazdu, wznowienie po przerwaniu,
// uzgadnianie przejazdu z sasiadem, tryb reczny.
//
// -------------------------------------------------------------
// SZEW DLA KLAS POCHODNYCH
// -------------------------------------------------------------
// Klasa pochodna w swoim ciele:
//   1. wypelnia wejscia czujnikow i napedu,
//   2. wola SUPER^(),
//   3. przepisuje xDrvRun / xDrvRev / lrDrvFreq na swoj aktuator.
//
// Dzieki temu logika sekwencji jest napisana RAZ i nie zalezy
// od tego, czy wezel ma napedy rolkowe, lancuchowe czy zadne.
//
// -------------------------------------------------------------
// DIAGNOSTYKA
// -------------------------------------------------------------
// Jesli wezel stoi, eWait mowi DOKLADNIE jednej rzeczy brakuje.
// Warunki sa sprawdzane w stalej kolejnosci i pierwszy
// niespelniony konczy cykl. Nie ma zagniezdzonych warunkow,
// w ktorych "cos" moze byc nie tak.
//
// -------------------------------------------------------------
// KONWENCJA ZAJETOSCI
// -------------------------------------------------------------
// Mem.xLoadPresent ustawiamy w chwili ROZPOCZECIA wjazdu, a
// kasujemy dopiero po potwierdzonym zjezdzie. W trakcie
// przejazdu oba wezly sa zajete - bo paleta fizycznie lezy
// na obu. To jest zalozenie bezpieczne: po zaniku zasilania
// wolimy jeden wezel za duzo do sprawdzenia niz kolizje.
VAR_INPUT

	// =========================================================
	// STEROWANIE NADRZEDNE
	// =========================================================

	eMode			: E_MachineMode;

	// TRUE = lancuch bezpieczenstwa zwolniony
	xSafetyOK		: BOOL;

	// Reczne zezwolenie na przejazdy miedzy stacjami.
	// FALSE zatrzymuje wydawanie ladunkow, nie ruszajac niczego
	// innego - sluzy do przechodzenia maszyny krok po kroku.
	xTransferEnable	: BOOL := TRUE;


	// =========================================================
	// SZEW CZUJNIKOW - wypelnia klasa pochodna PRZED SUPER^()
	// =========================================================

	// Przynajmniej jeden czujnik jest wlaczony przez operatora
	xSensUsable		: BOOL;

	// Ladunek w pozycji zatrzymania
	xSensLoadAtStop	: BOOL;

	// Pole czujnikow calkowicie wolne
	xSensLoadNone	: BOOL;

	// Czujniki nie zgadzaja sie ze soba
	xSensConflict	: BOOL;


	// =========================================================
	// SZEW NAPEDU - wypelnia klasa pochodna PRZED SUPER^()
	// =========================================================

	xDrvReady		: BOOL;
	xDrvFault		: BOOL;

END_VAR
VAR_OUTPUT

	// =========================================================
	// SZEW NAPEDU - czyta klasa pochodna PO SUPER^()
	// =========================================================

	xDrvRun			: BOOL;
	xDrvRev			: BOOL;
	lrDrvFreq		: LREAL;


	// =========================================================
	// DIAGNOSTYKA
	// =========================================================

	eState			: E_NodeState;

	// Jedyna przyczyna postoju w tym cyklu
	eWait			: E_WaitCause;

	eAlarm			: E_NodeAlarm;
	xAlarm			: BOOL;

	// Obraz z pamieci nieulotnej
	xOccupied		: BOOL;
	xLoadNok		: BOOL;

	// Operacja stacji zostala przerwana w polowie
	xOpInterrupted	: BOOL;

	// TRUE = pamiec sie zmienila, menedzer ma ja zapisac
	xPersistDirty	: BOOL;

END_VAR
VAR

	// Numer wezla - wylacznie do diagnostyki i HMI
	nNodeId			: INT;

	// Rekord nieulotny wezla - GVL_PERSIST.aConv[nNodeId]
	pP				: POINTER TO ST_ConvPersist;

	// Sasiedzi w lancuchu transportu
	pPrev			: POINTER TO FB_TransportNodeBase;
	pNext			: POINTER TO FB_TransportNodeBase;

	// Dokad przejsc po uplywie czasowki zatrzymania
	eStopTarget		: E_NodeState := NODE_OCCUPIED;

	eModeOld		: E_MachineMode;

	tonStopDelay	: TON;
	tonWatchdog		: TON;
	tonBlind		: TON;
	tonClear		: TON;
	tonSettle		: TON;

	xManFwd			: BOOL;
	xManRev			: BOOL;

END_VAR

// =============================================================
// CYKL WEZLA
// =============================================================
//
// Kolejnosc warunkow jest czescia specyfikacji - nie zmieniac
// bez zastanowienia. Pierwszy niespelniony warunek konczy cykl
// i zostaje w eWait jako jednoznaczna przyczyna postoju.


// -------------------------------------------------------------
// 1. KONFIGURACJA
// -------------------------------------------------------------

IF pP = 0 THEN
	M_HaltMotion();
	eWait	:= WAIT_NOT_CONFIGURED;
	eAlarm	:= ALM_NOT_CONFIGURED;
	xAlarm	:= TRUE;
	eState	:= NODE_ALARM;
	RETURN;
END_IF

xOccupied		:= pP^.Mem.xLoadPresent;
xLoadNok		:= pP^.Mem.xLoadNok;
xOpInterrupted	:= pP^.Mem.xOperationInterrupted;
xAlarm			:= (eAlarm <> ALM_NONE);


// -------------------------------------------------------------
// 2. BLAD NAPEDU
// -------------------------------------------------------------

IF xDrvFault THEN
	M_MarkAborted();
	M_RaiseAlarm(eNew := ALM_DRIVE_FAULT);
END_IF


// -------------------------------------------------------------
// 3. ZEZWOLENIE BEZPIECZENSTWA
// -------------------------------------------------------------
//
// Zanik STO w trakcie przejazdu zapamietujemy jako przerwany
// ruch. Po resecie maszyna sprobuje go dokonczyc sama.

IF NOT xSafetyOK THEN
	M_MarkAborted();
	M_MarkOperationInterrupted();
	M_HaltMotion();
	eWait := WAIT_NO_SAFETY;
	RETURN;
END_IF


// -------------------------------------------------------------
// 4. TRYB RECZNY
// -------------------------------------------------------------

IF eMode = MODE_MANUAL THEN
	eModeOld := eMode;
	M_ManualCycle();
	RETURN;
END_IF

IF eModeOld = MODE_MANUAL THEN
	// Po recznej maszyna nie wie, gdzie sa palety - weryfikujemy
	eState := NODE_INIT;
END_IF

eModeOld := eMode;


// -------------------------------------------------------------
// 5. ALARM
// -------------------------------------------------------------

IF xAlarm THEN
	M_HaltMotion();
	eWait	:= WAIT_ALARM_ACTIVE;
	eState	:= NODE_ALARM;
	RETURN;
END_IF


// -------------------------------------------------------------
// 6. PAMIEC NIEPOTWIERDZONA
// -------------------------------------------------------------
//
// Rozjazd pamieci z czujnikami rozstrzyga operator -
// M_ServiceSetEmpty albo M_ServiceSetLoaded.

IF NOT pP^.Mem.xStateVerified THEN
	M_HaltMotion();
	eWait	:= WAIT_STATE_UNVERIFIED;
	eState	:= NODE_VERIFY;
	RETURN;
END_IF


// -------------------------------------------------------------
// 7. TRYB INNY NIZ AUTO
// -------------------------------------------------------------

IF eMode <> MODE_AUTO THEN
	M_HaltMotion();
	eWait := WAIT_NOT_AUTO;
	RETURN;
END_IF


// -------------------------------------------------------------
// 8. SEKWENCJA AUTOMATYCZNA
// -------------------------------------------------------------

eWait := WAIT_NONE;

CASE eState OF

NODE_INIT:
	M_HaltMotion();
	M_CheckConsistency();

	IF NOT pP^.Mem.xStateVerified THEN
		RETURN;
	END_IF

	IF NOT pP^.Mem.xLoadPresent THEN
		eState := NODE_EMPTY;
		RETURN;
	END_IF

	// Ladunek lezy, ale operacja stacji nie zostala dokonczona -
	// wznawiamy ja zamiast wypuszczac nieprzebadana palete jako
	// dobra. Tu wraca maszyna po zaniku zasilania w polowie testu.
	IF M_OperationRequired() AND NOT pP^.Mem.xOperationDone THEN
		pP^.Mem.xOperationInterrupted	:= TRUE;
		xPersistDirty					:= TRUE;
		eState							:= NODE_BUSY;
		RETURN;
	END_IF

	eState := NODE_OCCUPIED;


NODE_EMPTY:
	M_HaltMotion();
	eWait := WAIT_NO_LOAD;
	M_CheckConsistency();


NODE_INFEED:
	M_RunForward();
	M_CheckInfeedWatchdog();

	// Hak dla stacji, ktore pracuja NA JADACEJ palecie -
	// stacja 4 dociska deski w trakcie przejazdu, stacja 6
	// skanuje profilometrem. Ich test konczy sie w chwili
	// dojazdu do czujnikow, a nie zaczyna po zatrzymaniu.
	M_TravelCycle();

	IF M_ArrivalDetected() THEN
		M_OnArrival();
	END_IF


NODE_STOP_DELAY:
	// Ladunek jest juz w pozycji, jedziemy jeszcze przez
	// czasowke ustawiona przez operatora
	M_RunForward();

	tonStopDelay(IN := TRUE, PT := pP^.Cfg.tStopDelay);

	IF tonStopDelay.Q THEN
		M_HaltMotion();
		M_ResetTravelTimers();

		pP^.Mem.xTransferAborted	:= FALSE;
		pP^.Mem.nResumeCount		:= 0;
		xPersistDirty				:= TRUE;

		eState := eStopTarget;
	END_IF


NODE_BUSY:
	M_HaltMotion();
	eWait := WAIT_OPERATION_BUSY;

	// Test przerwany na stacji, ktorej wyniku nie da sie
	// powtorzyc - paleta idzie na odrzut i nie jest juz badana
	IF pP^.Mem.xOperationInterrupted AND pP^.Cfg.xNokOnInterrupt THEN
		pP^.Mem.xLoadNok	:= TRUE;
		xPersistDirty		:= TRUE;
	END_IF

	IF M_OperationCycle() THEN
		pP^.Mem.xOperationDone	:= TRUE;
		xPersistDirty			:= TRUE;
		eState					:= NODE_OCCUPIED;
	END_IF


NODE_OCCUPIED:
	M_HaltMotion();
	M_CheckConsistency();

	IF eState = NODE_OCCUPIED THEN
		M_TryRelease();
	END_IF


NODE_OUTFEED:
	M_RunForward();
	M_CheckOutfeedWatchdog();

	IF M_ClearanceDetected() THEN
		M_OnCleared();
	END_IF


NODE_VERIFY:
	M_HaltMotion();
	eWait := WAIT_STATE_UNVERIFIED;


NODE_ALARM:
	M_HaltMotion();
	eWait := WAIT_ALARM_ACTIVE;


ELSE
	eState := NODE_INIT;

END_CASE


xOccupied		:= pP^.Mem.xLoadPresent;
xLoadNok		:= pP^.Mem.xLoadNok;
xOpInterrupted	:= pP^.Mem.xOperationInterrupted;
xAlarm			:= (eAlarm <> ALM_NONE);

METHOD PUBLIC M_Config
// Podpiecie rekordu nieulotnego. Wolac raz, przy starcie.
VAR_INPUT
	nId			: INT;
	pPersist	: POINTER TO ST_ConvPersist;
END_VAR
nNodeId	:= nId;
pP		:= pPersist;
END_METHOD

METHOD PUBLIC M_Link
// Podpiecie sasiadow w lancuchu transportu. Wolac raz.
VAR_INPUT
	pPrevNode	: POINTER TO FB_TransportNodeBase;
	pNextNode	: POINTER TO FB_TransportNodeBase;
END_VAR
pPrev := pPrevNode;
pNext := pNextNode;
END_METHOD

METHOD PUBLIC M_SetNext
// Zmiana nastepnika w trakcie pracy. Uzywa tego stacja
// rozjazdowa (8), ktora kieruje palete albo na sztaplarke,
// albo na transporter poprzeczny odrzutu.
VAR_INPUT
	pNextNode	: POINTER TO FB_TransportNodeBase;
END_VAR
pNext := pNextNode;
END_METHOD

METHOD PUBLIC M_ManJog
// Komendy ruchu recznego. Dzialaja tylko w MODE_MANUAL.
VAR_INPUT
	xFwd	: BOOL;
	xRev	: BOOL;
END_VAR
xManFwd := xFwd;
xManRev := xRev;
END_METHOD

METHOD PUBLIC M_Reset : BOOL
// Reset maszyny przez operatora.
//
// Jesli przejazd zostal przerwany (STO, zanik zasilania,
// watchdog), maszyna sama probuje go dokonczyc - wraca do
// fazy, w ktorej stanela, i ponawia ruch. Liczba prob jest
// nastawa operatora (nResumeRetries).
//
// Reset NIE potwierdza stanu pamieci. Jesli pamiec rozjechala
// sie z czujnikami, decyzje podejmuje operator przyciskiem
// "wezel pusty" albo "wezel zajety".
M_Reset := FALSE;

IF pP = 0 THEN
	RETURN;
END_IF


// ---------------------------------------------------------
// PRZERWANY PRZEJAZD - PROBA AUTOMATYCZNEGO DOKONCZENIA
// ---------------------------------------------------------

IF pP^.Mem.xTransferAborted THEN

	IF pP^.Mem.nResumeCount < pP^.Cfg.nResumeRetries THEN

		pP^.Mem.nResumeCount	:= pP^.Mem.nResumeCount + 1;
		xPersistDirty			:= TRUE;

		eAlarm	:= ALM_NONE;
		xAlarm	:= FALSE;

		M_ResetTravelTimers();

		eState	:= pP^.Mem.eAbortedPhase;
		M_Reset	:= TRUE;
		RETURN;

	END_IF

	// Proby wyczerpane - dalej decyduje czlowiek
	pP^.Mem.xStateVerified	:= FALSE;
	xPersistDirty			:= TRUE;

	eAlarm	:= ALM_RESUME_FAILED;
	xAlarm	:= TRUE;
	eState	:= NODE_VERIFY;
	RETURN;

END_IF


// ---------------------------------------------------------
// ZWYKLE KASOWANIE ALARMU
// ---------------------------------------------------------

eAlarm	:= ALM_NONE;
xAlarm	:= FALSE;

M_ResetTravelTimers();

eState	:= NODE_INIT;
M_Reset	:= TRUE;
END_METHOD

METHOD PUBLIC M_ServiceSetEmpty : BOOL
// Awaryjne kasowanie stanu.
//
// Serwis fizycznie zabral palete albo stos i potwierdza
// przyciskiem, ze wezel jest pusty. Kasuje pamiec, alarm
// i flage przerwanego przejazdu.
M_ServiceSetEmpty := FALSE;

IF pP = 0 THEN
	RETURN;
END_IF

pP^.Mem.xLoadPresent		:= FALSE;
pP^.Mem.xLoadNok			:= FALSE;
pP^.Mem.nLoadId				:= 0;
pP^.Mem.xOperationDone		:= FALSE;
pP^.Mem.xOperationInterrupted	:= FALSE;
pP^.Mem.xTransferAborted	:= FALSE;
pP^.Mem.nResumeCount		:= 0;
pP^.Mem.xStateVerified		:= TRUE;
xPersistDirty				:= TRUE;

eAlarm	:= ALM_NONE;
xAlarm	:= FALSE;

M_ResetTravelTimers();

eState				:= NODE_INIT;
M_ServiceSetEmpty	:= TRUE;
END_METHOD

METHOD PUBLIC M_ServiceSetLoaded : BOOL
// Operator potwierdza, ze na wezle LEZY ladunek i podaje
// jego werdykt. Uzywane, gdy czujnik padl albo gdy paleta
// zostala dolozona recznie.
VAR_INPUT
	xNok	: BOOL;
END_VAR
M_ServiceSetLoaded := FALSE;

IF pP = 0 THEN
	RETURN;
END_IF

pP^.Mem.xLoadPresent		:= TRUE;
pP^.Mem.xLoadNok			:= xNok;
// Paleta dolozona recznie nie byla badana - stacja ma to zrobic
pP^.Mem.xOperationDone		:= FALSE;
pP^.Mem.xOperationInterrupted	:= FALSE;
pP^.Mem.xTransferAborted	:= FALSE;
pP^.Mem.nResumeCount		:= 0;
pP^.Mem.xStateVerified		:= TRUE;
xPersistDirty				:= TRUE;

eAlarm	:= ALM_NONE;
xAlarm	:= FALSE;

M_ResetTravelTimers();

eState				:= NODE_INIT;
M_ServiceSetLoaded	:= TRUE;
END_METHOD

METHOD PUBLIC M_InjectLoad : BOOL
// Ladunek pojawia sie na wezle INNA droga niz transporterem.
//
// Operator wstawia stos na stacji 1, desztaplarka wydaje
// pojedyncza palete spod uniesionego stosu. W obu przypadkach
// nie bylo zadnego przejazdu, wiec wezel od razu przechodzi
// w stan zajety.
VAR_INPUT
	xNok	: BOOL;
	nLoadId	: UDINT;

	// TRUE = stacja ma juz ten ladunek obsluzony i moze go
	// wydac bez dalszej operacji
	xOpDone	: BOOL;
END_VAR
M_InjectLoad := FALSE;

IF pP = 0 THEN
	RETURN;
END_IF

pP^.Mem.xLoadPresent			:= TRUE;
pP^.Mem.xLoadNok				:= xNok;
pP^.Mem.nLoadId					:= nLoadId;
pP^.Mem.xOperationDone			:= xOpDone;
pP^.Mem.xOperationInterrupted	:= FALSE;
pP^.Mem.xTransferAborted		:= FALSE;
pP^.Mem.nResumeCount			:= 0;
pP^.Mem.xStateVerified			:= TRUE;
xPersistDirty					:= TRUE;

M_ResetTravelTimers();

eState			:= NODE_OCCUPIED;
M_InjectLoad	:= TRUE;
END_METHOD

METHOD PUBLIC M_ClearLoad : BOOL
// Ladunek opuscil wezel INNA droga niz transporterem -
// sztaplarka zabrala palete w gore, na szczeki.
//
// Nie myl tego z M_ServiceSetEmpty: tam operator rozstrzyga
// niezgodnosc pamieci z czujnikami, tu maszyna wie, co zrobila.
M_ClearLoad := FALSE;

IF pP = 0 THEN
	RETURN;
END_IF

pP^.Mem.xLoadPresent			:= FALSE;
pP^.Mem.xLoadNok				:= FALSE;
pP^.Mem.nLoadId					:= 0;
pP^.Mem.xOperationDone			:= FALSE;
pP^.Mem.xOperationInterrupted	:= FALSE;
pP^.Mem.xTransferAborted		:= FALSE;
pP^.Mem.nResumeCount			:= 0;
xPersistDirty					:= TRUE;

M_HaltMotion();
M_ResetTravelTimers();

eState		:= NODE_EMPTY;
M_ClearLoad	:= TRUE;
END_METHOD

METHOD PUBLIC M_AckPersist
// Menedzer zapisu danych nieulotnych potwierdza zapis.
xPersistDirty := FALSE;
END_METHOD

METHOD PUBLIC M_CanAccept : BOOL
// Czy wezel moze przyjac ladunek. Pyta o to poprzednik.
M_CanAccept := (M_WhyCannotAccept() = WAIT_NONE);
END_METHOD

METHOD PUBLIC M_WhyCannotAccept : E_WaitCause
// Jedna, konkretna przyczyna odmowy przyjecia ladunku.
// Poprzednik przepisuje ja do swojego eWait, dzieki czemu
// na HMI widac nie "wezel czeka", tylko czego dokladnie
// brakuje i po ktorej stronie.
M_WhyCannotAccept := WAIT_NONE;

IF pP = 0 THEN
	M_WhyCannotAccept := WAIT_NOT_CONFIGURED;
	RETURN;
END_IF

IF NOT xSafetyOK THEN
	M_WhyCannotAccept := WAIT_NEXT_NO_SAFETY;
	RETURN;
END_IF

IF eMode <> MODE_AUTO THEN
	M_WhyCannotAccept := WAIT_NEXT_NOT_AUTO;
	RETURN;
END_IF

IF eAlarm <> ALM_NONE THEN
	M_WhyCannotAccept := WAIT_NEXT_ALARM;
	RETURN;
END_IF

IF NOT pP^.Mem.xStateVerified THEN
	M_WhyCannotAccept := WAIT_NEXT_UNVERIFIED;
	RETURN;
END_IF

IF pP^.Mem.xLoadPresent THEN
	M_WhyCannotAccept := WAIT_NEXT_OCCUPIED;
	RETURN;
END_IF

IF eState = NODE_BUSY THEN
	M_WhyCannotAccept := WAIT_NEXT_BUSY;
	RETURN;
END_IF

IF eState <> NODE_EMPTY THEN
	M_WhyCannotAccept := WAIT_NEXT_OCCUPIED;
	RETURN;
END_IF
END_METHOD

METHOD PUBLIC M_RequiresPrevStop : BOOL
// Czy poprzednik MUSI zatrzymac ladunek u siebie.
//
// Wezel z wylaczonymi oboma czujnikami mierzy przejazd
// czasowka. Zeby ten czas cokolwiek znaczyl, ladunek musi
// ruszac zawsze z tego samego miejsca - wiec poprzednik
// nie ma prawa przepuscic go bez zatrzymania.
IF pP = 0 THEN
	M_RequiresPrevStop := TRUE;
	RETURN;
END_IF

M_RequiresPrevStop := NOT (pP^.Cfg.xSensor1Enabled OR pP^.Cfg.xSensor2Enabled);
END_METHOD

METHOD PUBLIC M_BeginInfeed
// Poprzednik zaczyna wydawanie. Oba wezly rusza w tym samym
// cyklu - ten przechodzi na NODE_INFEED, tamten na NODE_OUTFEED.
VAR_INPUT
	pSource		: POINTER TO FB_TransportNodeBase;
	xNok		: BOOL;
	nLoadId		: UDINT;
END_VAR
IF pP = 0 THEN
	RETURN;
END_IF

pPrev := pSource;

// Zajetosc ustawiamy JUZ TERAZ - paleta wchodzi na wezel
pP^.Mem.xLoadPresent		:= TRUE;
pP^.Mem.xLoadNok			:= xNok;
pP^.Mem.nLoadId				:= nLoadId;
pP^.Mem.xOperationDone		:= FALSE;
pP^.Mem.xOperationInterrupted	:= FALSE;
pP^.Mem.xTransferAborted	:= FALSE;
pP^.Mem.nResumeCount		:= 0;
xPersistDirty				:= TRUE;

M_ResetTravelTimers();

eState := NODE_INFEED;
END_METHOD

METHOD PROTECTED M_TryRelease : BOOL
// Proba wydania ladunku dalej. Jesli nastepnik jest gotowy,
// oba transportery rusza w tym samym cyklu.
M_TryRelease := FALSE;

IF NOT xTransferEnable THEN
	eWait := WAIT_TRANSFER_HOLD;
	RETURN;
END_IF

IF pNext = 0 THEN
	eWait := WAIT_NEXT_NOT_LINKED;
	RETURN;
END_IF

eWait := pNext^.M_WhyCannotAccept();

IF eWait <> WAIT_NONE THEN
	RETURN;
END_IF

pNext^.M_BeginInfeed(
	pSource	:= ADR(THIS^),
	xNok	:= pP^.Mem.xLoadNok,
	nLoadId	:= pP^.Mem.nLoadId
);

M_ResetTravelTimers();

eState			:= NODE_OUTFEED;
M_TryRelease	:= TRUE;
END_METHOD

METHOD PROTECTED M_PassThroughPossible : BOOL
// Czy mozna przepuscic ladunek bez zatrzymania.
//
// Sens: jesli na tym wezle nie ma nic do zrobienia, a
// nastepny czeka na palete, to zatrzymywanie jej tutaj
// tylko traci czas i zuzywa maszyne.
M_PassThroughPossible := FALSE;

IF NOT pP^.Cfg.xAllowPassThrough THEN
	RETURN;
END_IF

IF pNext = 0 THEN
	RETURN;
END_IF

// Nastepnik jedzie na czasowke - potrzebuje powtarzalnego
// punktu startu, wiec musimy zatrzymac palete u siebie
IF pNext^.M_RequiresPrevStop() THEN
	RETURN;
END_IF

IF NOT pNext^.M_CanAccept() THEN
	RETURN;
END_IF

M_PassThroughPossible := TRUE;
END_METHOD

METHOD PROTECTED M_OnArrival
// Ladunek dojechal do pozycji koncowej. Trzy mozliwosci,
// sprawdzane w tej kolejnosci.
M_ResetTravelTimers();


// 1. Stacja ma cos do zrobienia - zatrzymujemy zawsze
IF M_OperationRequired() THEN
	eStopTarget	:= NODE_BUSY;
	eState		:= NODE_STOP_DELAY;
	RETURN;
END_IF


// 2. Nie ma nic do zrobienia, nastepnik czeka - jedziemy dalej
IF M_PassThroughPossible() THEN
	IF M_TryRelease() THEN
		RETURN;
	END_IF
END_IF


// 3. Zatrzymanie w pozycji koncowej
eStopTarget	:= NODE_OCCUPIED;
eState		:= NODE_STOP_DELAY;
END_METHOD

METHOD PROTECTED M_OnCleared
// Ladunek potwierdzenie zjechal z wezla.
pP^.Mem.xLoadPresent		:= FALSE;
pP^.Mem.xLoadNok			:= FALSE;
pP^.Mem.nLoadId				:= 0;
pP^.Mem.xOperationDone		:= FALSE;
pP^.Mem.xOperationInterrupted	:= FALSE;
pP^.Mem.xTransferAborted	:= FALSE;
pP^.Mem.nResumeCount		:= 0;
xPersistDirty				:= TRUE;

M_HaltMotion();
M_ResetTravelTimers();

eState := NODE_EMPTY;
END_METHOD

METHOD PROTECTED M_ArrivalDetected : BOOL
// Wykrycie pozycji koncowej. Przy wylaczonych obu czujnikach
// zastepuje je czasowka nastawiana przez operatora.
IF xSensUsable THEN
	tonBlind(IN := FALSE);
	M_ArrivalDetected := xSensLoadAtStop;
	RETURN;
END_IF

tonBlind(IN := TRUE, PT := pP^.Cfg.tBlindTravel);
M_ArrivalDetected := tonBlind.Q;
END_METHOD

METHOD PROTECTED M_ClearanceDetected : BOOL
// Potwierdzenie, ze ladunek zszedl z pola czujnikow.
VAR
	xFree	: BOOL;
END_VAR
IF xSensUsable THEN
	tonBlind(IN := FALSE);
	xFree := xSensLoadNone;
ELSE
	tonBlind(IN := TRUE, PT := pP^.Cfg.tBlindTravel);
	xFree := tonBlind.Q;
END_IF

tonClear(IN := xFree, PT := pP^.Cfg.tClearDelay);

M_ClearanceDetected := tonClear.Q;
END_METHOD

METHOD PROTECTED M_CheckInfeedWatchdog
// Paleta miala dojechac i nie dojechala - zaciecie, poslizg,
// urwany lancuch. Zatrzymujemy i wolamy operatora.
tonWatchdog(IN := TRUE, PT := pP^.Cfg.tInfeedWatchdog);

IF NOT tonWatchdog.Q THEN
	RETURN;
END_IF

M_MarkAborted();
M_RaiseAlarm(eNew := ALM_INFEED_TIMEOUT);
eState := NODE_ALARM;
END_METHOD

METHOD PROTECTED M_CheckOutfeedWatchdog
// Paleta miala zjechac i nie zjechala.
tonWatchdog(IN := TRUE, PT := pP^.Cfg.tOutfeedWatchdog);

IF NOT tonWatchdog.Q THEN
	RETURN;
END_IF

M_MarkAborted();
M_RaiseAlarm(eNew := ALM_OUTFEED_TIMEOUT);
eState := NODE_ALARM;
END_METHOD

METHOD PROTECTED M_CheckConsistency
// Weryfikacja pamieci wzgledem czujnikow. Wolana na postoju:
// po zatrzymaniu, w stanie pustym i przy starcie.
//
// Niezgodnosc musi utrzymac sie przez tSensorSettle, zeby nie
// lapac drgan i kostek palety migajacych czujnikowi.
VAR
	eDetect	: E_NodeAlarm;
END_VAR
IF NOT xSensUsable THEN
	tonSettle(IN := FALSE);
	RETURN;
END_IF

// Stacje, ktore zdejmuja ladunek z transportera wlasna mechanika
// (desztaplarka, sztaplarka), wstrzymuja to porownanie na czas
// swojego cyklu - patrz M_SensorCheckAllowed.
IF NOT M_SensorCheckAllowed() THEN
	tonSettle(IN := FALSE);
	RETURN;
END_IF

eDetect := ALM_NONE;

IF pP^.Mem.xLoadPresent THEN

	IF xSensLoadNone THEN
		// Pamiec mowi "zajete", czujniki nie widza nic
		eDetect := ALM_LOAD_LOST;
	ELSIF xSensConflict THEN
		// Jeden czujnik widzi, drugi nie - paleta krzywo
		// albo czujnik padl
		eDetect := ALM_SENSOR_DISAGREE;
	END_IF

ELSE

	IF NOT xSensLoadNone THEN
		// Pamiec mowi "pusto", a cos tam lezy
		eDetect := ALM_UNEXPECTED_LOAD;
	END_IF

END_IF


tonSettle(IN := (eDetect <> ALM_NONE), PT := pP^.Cfg.tSensorSettle);

IF NOT tonSettle.Q THEN
	RETURN;
END_IF

pP^.Mem.xStateVerified	:= FALSE;
xPersistDirty			:= TRUE;

M_RaiseAlarm(eNew := eDetect);
eState := NODE_VERIFY;
END_METHOD

METHOD PROTECTED M_MarkAborted
// Zapamietanie, ze ruch zostal przerwany w polowie. Po
// resecie maszyna wroci dokladnie do tej fazy i sprobuje
// dokonczyc przejazd.
IF pP = 0 THEN
	RETURN;
END_IF

IF (eState <> NODE_INFEED) AND (eState <> NODE_OUTFEED) AND (eState <> NODE_STOP_DELAY) THEN
	RETURN;
END_IF

IF pP^.Mem.xTransferAborted THEN
	RETURN;
END_IF

pP^.Mem.xTransferAborted	:= TRUE;
pP^.Mem.eAbortedPhase		:= eState;
xPersistDirty				:= TRUE;
END_METHOD

METHOD PROTECTED M_MarkOperationInterrupted
// Operacja stacji zostala przerwana w polowie.
//
// Sama flaga nie przesadza o losie palety - o tym decyduje
// Cfg.xNokOnInterrupt. Na stacjach 4 i 6 wyniku przerwanego
// testu nie da sie uznac za wiarygodny, wiec paleta idzie na
// odrzut. Na pozostalych mozna kontynuowac albo powtorzyc cykl.
IF pP = 0 THEN
	RETURN;
END_IF

IF eState <> NODE_BUSY THEN
	RETURN;
END_IF

IF pP^.Mem.xOperationInterrupted THEN
	RETURN;
END_IF

pP^.Mem.xOperationInterrupted	:= TRUE;
xPersistDirty					:= TRUE;
END_METHOD

METHOD PROTECTED M_RaiseAlarm
// Pierwszy alarm zostaje - kolejne go nie nadpisza, zeby
// operator widzial przyczyne, a nie skutek.
VAR_INPUT
	eNew	: E_NodeAlarm;
END_VAR
IF eNew = ALM_NONE THEN
	RETURN;
END_IF

IF eAlarm = ALM_NONE THEN
	eAlarm := eNew;
END_IF

xAlarm := TRUE;

// Alarm w trakcie operacji to przerwanie testu - grzyb,
// kurtyna, przeciazenie napedu. Na stacjach 4 i 6 unieważnia
// wynik, na pozostalych tylko wstrzymuje cykl.
M_MarkOperationInterrupted();

M_HaltMotion();
END_METHOD

METHOD PROTECTED M_HaltMotion
xDrvRun		:= FALSE;
xDrvRev		:= FALSE;
lrDrvFreq	:= 0.0;
END_METHOD

METHOD PROTECTED M_RunForward
// W AUTO transporter jedzie zawsze do przodu.
xDrvRun		:= TRUE;
xDrvRev		:= FALSE;
lrDrvFreq	:= pP^.Cfg.lrFreqAuto;
END_METHOD

METHOD PROTECTED M_ResetTravelTimers
tonWatchdog(IN := FALSE);
tonBlind(IN := FALSE);
tonClear(IN := FALSE);
tonStopDelay(IN := FALSE);
tonSettle(IN := FALSE);
END_METHOD

METHOD PROTECTED M_ManualCycle
// Praca reczna: ruch w obie strony, bez uzgadniania z
// sasiadami i bez watchdogow. Pamiec obecnosci NIE jest
// aktualizowana - po powrocie do AUTO wezel przechodzi
// przez NODE_INIT i weryfikuje stan czujnikami.
eState	:= NODE_MANUAL;
eWait	:= WAIT_NONE;

M_ResetTravelTimers();

IF xManFwd AND NOT xManRev THEN
	xDrvRun		:= TRUE;
	xDrvRev		:= FALSE;
	lrDrvFreq	:= pP^.Cfg.lrFreqManual;
	RETURN;
END_IF

IF xManRev AND NOT xManFwd THEN
	xDrvRun		:= TRUE;
	xDrvRev		:= TRUE;
	lrDrvFreq	:= pP^.Cfg.lrFreqManual;
	RETURN;
END_IF

M_HaltMotion();
END_METHOD

METHOD PROTECTED M_OperationRequired : BOOL
// HAK DLA STACJI TECHNOLOGICZNYCH.
//
// TRUE = paleta musi sie tu zatrzymac, bo jest co robic.
// Klasa pochodna nadpisuje i uwzglednia:
//   - Cfg.xStationEnabled (operator wylaczyl stacje),
//   - Mem.xLoadNok (paleta odrzucona - zadnych dalszych testow).
//
// Domyslnie wezel jest samym transporterem.
M_OperationRequired := FALSE;
END_METHOD

METHOD PROTECTED M_SensorCheckAllowed : BOOL
// HAK DLA STACJI Z WLASNA MECHANIKA NAD TRANSPORTEREM.
//
// FALSE wstrzymuje porownanie pamieci z czujnikami. Potrzebuja
// tego desztaplarka i sztaplarka: u nich stos potrafi wisiec na
// szczekach albo schodzic na transporter w chwili, gdy pamiec
// wezla mowi "pusto", i odwrotnie.
//
// Domyslnie TRUE - zwykly transporter porownuje zawsze.
M_SensorCheckAllowed := TRUE;
END_METHOD

METHOD PROTECTED M_TravelCycle
// HAK DLA STACJI PRACUJACYCH NA JADACEJ PALECIE.
//
// Wolany w kazdym cyklu, gdy ladunek wjezdza na wezel.
//
// Stacja 4 dociska deski rolkami w trakcie przejazdu, stacja 6
// skanuje profilometrem milimetr po milimetrze. Dla nich test
// nie zaczyna sie po zatrzymaniu - on trwa CALY przejazd
// i konczy sie w chwili dojazdu do czujnikow.
//
// Wlasnie dlatego przerwanie na tych stacjach uniewaznia wynik:
// paleta zatrzymuje sie w nieznanym miejscu, a po wznowieniu
// nie da sie odtworzyc warunkow, w ktorych badanie sie toczylo.
//
// Domyslnie pusty - zwykly transporter nic po drodze nie robi.
;
END_METHOD

METHOD PROTECTED M_OperationCycle : BOOL
// HAK DLA STACJI TECHNOLOGICZNYCH.
// TRUE = operacja zakonczona, paleta moze jechac dalej.
M_OperationCycle := TRUE;
END_METHOD

END_FUNCTION_BLOCK

// ---- POUs/POUs/FB/FB_Station11_Stack.TcPOU
FUNCTION_BLOCK FB_Station11_Stack EXTENDS FB_RollerConveyor
// =============================================================
// STACJA 11 - SZTAPLARKA
// =============================================================
//
// Ta sama kinematyka co desztaplarka, sekwencja odwrocona.
// Wozek trzyma rosnacy stos w gorze, a kazda nowa paleta
// wjezdza pod niego.
//
// -------------------------------------------------------------
// CYKL
// -------------------------------------------------------------
//   czekanie      wozek na GORZE, szczeki zamkniete na stosie
//   wjazd palety  paleta zatrzymuje sie na czujnikach
//   odlozenie     wozek na SRODEK - stos siada na nowa palete
//   otwarcie      szczeki puszczaja stos
//   zejscie       wozek na DOL, pod najnizsza palete
//   chwyt         szczeki zamykaja sie na calym stosie
//   uniesienie    wozek na GORE, stos wyzszy o jedna palete
//   i od nowa, az uzbiera sie Cfg.nStackSize sztuk
//
// -------------------------------------------------------------
// KOLIZJA
// -------------------------------------------------------------
// Paleta nie ma prawa wjechac, dopoki wozek nie stoi na GORZE
// z zamknietymi szczekami. Inaczej wjechalaby wprost w stos
// albo w szczeki - dlatego jest to warunek przyjecia ladunku,
// a nie tylko krok sekwencji.
VAR_INPUT

	diLiftPosRaw	: DINT;
	xJawClosedSw	: BOOL;
	xJawOpenSw		: BOOL;

END_VAR
VAR_OUTPUT

	xJawCoilClose	: BOOL;
	xJawCoilOpen	: BOOL;

	nStep			: INT;

	// Ile palet wisi na szczekach
	nHeld			: INT;

	diLiftPos		: DINT;
	nLiftTarget		: INT;
	xLiftInPos		: BOOL;

	eLiftAlarm		: E_StackAlarm;

END_VAR
VAR

	pSt		: POINTER TO ST_StackPersist;
	fbLift	: FB_StackLift;

	nStackId	: UDINT;

END_VAR
VAR CONSTANT

	ST11_IDLE		: INT := 0;
	ST11_SETDOWN	: INT := 10;
	ST11_OPEN		: INT := 20;
	ST11_GODOWN		: INT := 30;
	ST11_GRIP		: INT := 40;
	ST11_LIFT		: INT := 50;
	ST11_AFTER		: INT := 60;
	ST11_DELIVER	: INT := 70;
	ST11_RELEASE	: INT := 80;

END_VAR

// =============================================================
// CYKL STACJI 11
// =============================================================


M_CallLift();

SUPER^();

M_StackCycle();

M_MapStatus();

METHOD PUBLIC M_ConfigStation
// Wolac raz, przy starcie, PO M_Config klasy bazowej.
VAR_INPUT
	pStPersist	: POINTER TO ST_StackPersist;

	// Falownik krzywki sztaplarki
	pLiftDrive	: POINTER TO FB_NordSK550PP;

	nJawId		: INT;
	pJawPersist	: POINTER TO ST_CylPersist;
END_VAR
pSt := pStPersist;

fbLift.M_Config(
	pPersist	:= pStPersist,
	pDrv		:= pLiftDrive,
	nJawId		:= nJawId,
	pJawPersist	:= pJawPersist
);
END_METHOD

METHOD PROTECTED M_CallLift
fbLift(
	eMode			:= eMode,
	xSafetyOK		:= xSafetyOK,
	diPosRaw		:= diLiftPosRaw,
	xJawClosedSw	:= xJawClosedSw,
	xJawOpenSw		:= xJawOpenSw
);

xJawCoilClose	:= fbLift.xJawCoilClose;
xJawCoilOpen	:= fbLift.xJawCoilOpen;

IF fbLift.xAlarm THEN
	M_RaiseAlarm(eNew := ALM_OPERATION_FAILED);
END_IF
END_METHOD

METHOD PROTECTED M_MapStatus
diLiftPos	:= fbLift.diPos;
nLiftTarget	:= fbLift.nTargetSel;
xLiftInPos	:= fbLift.xInPosition;
eLiftAlarm	:= fbLift.eAlarm;

IF pSt <> 0 THEN
	nHeld := pSt^.Mem.nHeld;
END_IF
END_METHOD

METHOD PUBLIC M_WhyCannotAccept : E_WaitCause
// Warunki klasy bazowej plus zabezpieczenie przed kolizja:
// wozek musi stac na GORZE, a jesli cos trzyma - ze
// szczekami zamknietymi.
M_WhyCannotAccept := SUPER^.M_WhyCannotAccept();

IF M_WhyCannotAccept <> WAIT_NONE THEN
	RETURN;
END_IF

IF pSt = 0 THEN
	M_WhyCannotAccept := WAIT_NOT_CONFIGURED;
	RETURN;
END_IF

// Stacja wylaczona - sam przelot, bez warunkow mechaniki
IF NOT pP^.Cfg.xStationEnabled THEN
	RETURN;
END_IF

IF (fbLift.nTargetSel <> 3) OR NOT fbLift.xInPosition THEN
	M_WhyCannotAccept := WAIT_STATION_NOT_READY;
	RETURN;
END_IF

IF (pSt^.Mem.nHeld > 0) AND NOT fbLift.xJawsClosed THEN
	M_WhyCannotAccept := WAIT_STATION_NOT_READY;
END_IF
END_METHOD

METHOD PROTECTED M_OperationRequired : BOOL
// Kazda paleta musi sie zatrzymac i trafic na stos. Gotowy stos
// wydany przez M_InjectLoad ma juz xOperationDone.
M_OperationRequired := TRUE;

IF pP = 0 THEN
	RETURN;
END_IF

IF NOT pP^.Cfg.xStationEnabled THEN
	M_OperationRequired := FALSE;
	RETURN;
END_IF

M_OperationRequired := NOT pP^.Mem.xOperationDone;
END_METHOD

METHOD PROTECTED M_OperationCycle : BOOL
// Wlasciwa sekwencja siedzi w M_StackCycle - musi dzialac takze
// wtedy, gdy wezel jest pusty, bo wozek konczy wtedy ruch w gore.
M_OperationCycle := FALSE;

IF pP = 0 THEN
	RETURN;
END_IF

M_OperationCycle := pP^.Mem.xOperationDone;
END_METHOD

